(* IEC 61131-3 sources: TetherPLC/compat/tc2 (part 2) *)

(* ---- tc2_hvac.st ---- *)
// tc2_hvac.st — Tc2_HVAC surface (TF8000_TC3_HVAC_EN): pure-ST
// HVAC control blocks — no host/hardware dependency.  Covers
// the documented categories: actuators, motors/pumps, mux,
// redundancy, analog scaling, controllers (2-point, step, PID),
// sequence controllers, heating curve / outside-temp damping,
// alarm/anti-blocking/blink helpers, and BAR room-automation
// primitives.  Terminal bindings (KL32xx) are not modeled —
// the blocks operate on scaled process values.

// ---- FB_HVACAnalogInput: raw counts -> engineering value ----
FUNCTION_BLOCK FB_HVACAnalogInput
VAR_INPUT
    Raw : LREAL;                // raw counts
    RawMin : LREAL;
    RawMax : LREAL;
    EngMin : LREAL;
    EngMax : LREAL;
END_VAR
VAR_OUTPUT
    Value : LREAL;
END_VAR
    IF RawMax = RawMin THEN
        Value := EngMin;
    ELSE
        Value := EngMin + (Raw - RawMin) * (EngMax - EngMin) /
                 (RawMax - RawMin);
        IF Value < EngMin THEN Value := EngMin; END_IF;
        IF Value > EngMax THEN Value := EngMax; END_IF;
    END_IF;
END_FUNCTION_BLOCK

// ---- FB_HVACAnalogOutput: engineering value -> raw ----
FUNCTION_BLOCK FB_HVACAnalogOutput
VAR_INPUT
    Value : LREAL;
    EngMin : LREAL;
    EngMax : LREAL;
    RawMin : LREAL;
    RawMax : LREAL;
END_VAR
VAR_OUTPUT
    Raw : LREAL;
END_VAR
    IF EngMax = EngMin THEN
        Raw := RawMin;
    ELSE
        Raw := RawMin + (Value - EngMin) * (RawMax - RawMin) /
               (EngMax - EngMin);
        IF Raw < RawMin THEN Raw := RawMin; END_IF;
        IF Raw > RawMax THEN Raw := RawMax; END_IF;
    END_IF;
END_FUNCTION_BLOCK

// ---- FB_HVACScale: generic piecewise-linear scale ----
FUNCTION_BLOCK FB_HVACScale
VAR_INPUT
    x : LREAL;
    xMin : LREAL;
    xMax : LREAL;
    yMin : LREAL;
    yMax : LREAL;
END_VAR
VAR_OUTPUT
    y : LREAL;
END_VAR
    IF xMax = xMin THEN
        y := yMin;
    ELSE
        y := yMin + (x - xMin) * (yMax - yMin) / (xMax - xMin);
    END_IF;
END_FUNCTION_BLOCK

// ---- FB_HVAC2PointActuator: two-point damper/valve ----
// bCtrlVoltage TRUE -> run open; plus manual override and end-
// switch feedback monitoring.
FUNCTION_BLOCK FB_HVAC2PointActuator
VAR_INPUT
    bEnable : BOOL;
    bIn : BOOL;                 // demand: TRUE = open
    bManSwitch : BOOL;          // manual open override
    bLimitSwitchOpen : BOOL;
    bLimitSwitchClose : BOOL;
    tRun : LREAL;               // travel time s
    CycleTime : LREAL;
END_VAR
VAR_OUTPUT
    bOut : BOOL;                // drive command
    bFault : BOOL;              // end-switch disagreement
    Position : LREAL;           // 0 closed .. 100 open
END_VAR
VAR
    pos : LREAL;
END_VAR
    IF NOT bEnable THEN
        bOut := FALSE;
        bFault := FALSE;
        RETURN;
    END_IF;
    bOut := bIn OR bManSwitch;
    IF tRun > 0.0 THEN
        IF bOut THEN
            pos := pos + 100.0 * CycleTime / tRun;
            IF pos > 100.0 THEN pos := 100.0; END_IF;
        ELSE
            pos := pos - 100.0 * CycleTime / tRun;
            IF pos < 0.0 THEN pos := 0.0; END_IF;
        END_IF;
    END_IF;
    Position := pos;
    // fault: fully driven but feedback contradicts
    bFault := (pos >= 100.0 AND NOT bLimitSwitchOpen) OR
             (pos <= 0.0 AND NOT bLimitSwitchClose);
END_FUNCTION_BLOCK

// ---- FB_HVAC3PointActuator: three-point (open/close) ----
FUNCTION_BLOCK FB_HVAC3PointActuator
VAR_INPUT
    bEnable : BOOL;
    bOpen : BOOL;
    bClose : BOOL;
    tRun : LREAL;
    CycleTime : LREAL;
END_VAR
VAR_OUTPUT
    bOutOpen : BOOL;
    bOutClose : BOOL;
    Position : LREAL;
END_VAR
VAR
    pos : LREAL;
END_VAR
    IF NOT bEnable THEN
        bOutOpen := FALSE;
        bOutClose := FALSE;
        RETURN;
    END_IF;
    bOutOpen := bOpen AND NOT bClose;
    bOutClose := bClose AND NOT bOpen;
    IF tRun > 0.0 THEN
        IF bOutOpen THEN
            pos := pos + 100.0 * CycleTime / tRun;
            IF pos > 100.0 THEN pos := 100.0; END_IF;
        END_IF;
        IF bOutClose THEN
            pos := pos - 100.0 * CycleTime / tRun;
            IF pos < 0.0 THEN pos := 0.0; END_IF;
        END_IF;
    END_IF;
    Position := pos;
END_FUNCTION_BLOCK

// ---- FB_HVACCirculationPump: pump with standby lead swap ----
FUNCTION_BLOCK FB_HVACCirculationPump
VAR_INPUT
    bEnable : BOOL;
    bDemand : BOOL;
    bFault1 : BOOL;
    bFault2 : BOOL;
    bSwap : BOOL;               // lead-rotation request
END_VAR
VAR_OUTPUT
    bPump1 : BOOL;
    bPump2 : BOOL;
    Lead : INT;                 // 1 or 2
    bAlarm : BOOL;
END_VAR
VAR
    leadN : INT;
END_VAR
    IF leadN = 0 THEN leadN := 1; END_IF;
    IF bSwap THEN
        IF leadN = 1 THEN leadN := 2; ELSE leadN := 1; END_IF;
    END_IF;
    Lead := leadN;
    IF NOT bEnable OR NOT bDemand THEN
        bPump1 := FALSE;
        bPump2 := FALSE;
        bAlarm := bFault1 AND bFault2;
        RETURN;
    END_IF;
    bPump1 := leadN = 1 AND NOT bFault1;
    bPump2 := (leadN = 2 OR bFault1) AND NOT bFault2;
    bAlarm := bFault1 AND bFault2;
END_FUNCTION_BLOCK

// ---- FB_HVACMotor1Speed / Motor2Speed / Motor3Speed ----
FUNCTION_BLOCK FB_HVACMotor1Speed
VAR_INPUT
    bEnable : BOOL;
    Speed : INT;                // 0 off, 1 run
END_VAR
VAR_OUTPUT
    bOut1 : BOOL;
END_VAR
    bOut1 := bEnable AND Speed = 1;
END_FUNCTION_BLOCK

FUNCTION_BLOCK FB_HVACMotor2Speed
VAR_INPUT
    bEnable : BOOL;
    Speed : INT;                // 0..2
END_VAR
VAR_OUTPUT
    bOut1 : BOOL;
    bOut2 : BOOL;
END_VAR
    bOut1 := bEnable AND Speed = 1;
    bOut2 := bEnable AND Speed = 2;
END_FUNCTION_BLOCK

FUNCTION_BLOCK FB_HVACMotor3Speed
VAR_INPUT
    bEnable : BOOL;
    Speed : INT;                // 0..3
END_VAR
VAR_OUTPUT
    bOut1 : BOOL;
    bOut2 : BOOL;
    bOut3 : BOOL;
END_VAR
    bOut1 := bEnable AND Speed = 1;
    bOut2 := bEnable AND Speed = 2;
    bOut3 := bEnable AND Speed = 3;
END_FUNCTION_BLOCK

// ---- FB_HVACMux8: 8 -> 1 analog mux by selector ----
FUNCTION_BLOCK FB_HVACMux8
VAR_INPUT
    Sel : INT;                  // 1..8
    In1 : LREAL; In2 : LREAL; In3 : LREAL; In4 : LREAL;
    In5 : LREAL; In6 : LREAL; In7 : LREAL; In8 : LREAL;
END_VAR
VAR_OUTPUT
    Out : LREAL;
END_VAR
    IF Sel = 1 THEN Out := In1;
    ELSIF Sel = 2 THEN Out := In2;
    ELSIF Sel = 3 THEN Out := In3;
    ELSIF Sel = 4 THEN Out := In4;
    ELSIF Sel = 5 THEN Out := In5;
    ELSIF Sel = 6 THEN Out := In6;
    ELSIF Sel = 7 THEN Out := In7;
    ELSIF Sel = 8 THEN Out := In8;
    ELSE Out := 0.0;
    END_IF;
END_FUNCTION_BLOCK

// ---- FB_HVACMux8_BOOL: 8 -> 1 bool mux ----
FUNCTION_BLOCK FB_HVACMux8_BOOL
VAR_INPUT
    Sel : INT;
    In1 : BOOL; In2 : BOOL; In3 : BOOL; In4 : BOOL;
    In5 : BOOL; In6 : BOOL; In7 : BOOL; In8 : BOOL;
END_VAR
VAR_OUTPUT
    Out : BOOL;
END_VAR
    IF Sel = 1 THEN Out := In1;
    ELSIF Sel = 2 THEN Out := In2;
    ELSIF Sel = 3 THEN Out := In3;
    ELSIF Sel = 4 THEN Out := In4;
    ELSIF Sel = 5 THEN Out := In5;
    ELSIF Sel = 6 THEN Out := In6;
    ELSIF Sel = 7 THEN Out := In7;
    ELSIF Sel = 8 THEN Out := In8;
    ELSE Out := FALSE;
    END_IF;
END_FUNCTION_BLOCK

// ---- FB_HVACRedundancyCtrl: n+1 pump/fan redundancy ----
// N units, need Required running; rotates the lead and covers
// faults in order.
FUNCTION_BLOCK FB_HVACRedundancyCtrl
VAR_INPUT
    bEnable : BOOL;
    Required : INT;             // units demanded 0..3
    bFault1 : BOOL;
    bFault2 : BOOL;
    bFault3 : BOOL;
    bRotate : BOOL;
END_VAR
VAR_OUTPUT
    bOut1 : BOOL;
    bOut2 : BOOL;
    bOut3 : BOOL;
    Lead : INT;
    bAlarm : BOOL;
END_VAR
VAR
    leadN : INT;
    want : INT;
    ok1 : BOOL;
    ok2 : BOOL;
    ok3 : BOOL;
END_VAR
    IF leadN = 0 THEN leadN := 1; END_IF;
    IF bRotate THEN
        leadN := leadN + 1;
        IF leadN > 3 THEN leadN := 1; END_IF;
    END_IF;
    Lead := leadN;
    ok1 := NOT bFault1;
    ok2 := NOT bFault2;
    ok3 := NOT bFault3;
    want := Required;
    bOut1 := FALSE; bOut2 := FALSE; bOut3 := FALSE;
    IF bEnable THEN
        // start at leadN, wrap, pick healthy units
        IF want > 0 THEN
            IF leadN = 1 THEN
                IF ok1 THEN bOut1 := TRUE; want := want - 1; END_IF;
                IF want > 0 AND ok2 THEN bOut2 := TRUE; want := want - 1; END_IF;
                IF want > 0 AND ok3 THEN bOut3 := TRUE; want := want - 1; END_IF;
            ELSIF leadN = 2 THEN
                IF ok2 THEN bOut2 := TRUE; want := want - 1; END_IF;
                IF want > 0 AND ok3 THEN bOut3 := TRUE; want := want - 1; END_IF;
                IF want > 0 AND ok1 THEN bOut1 := TRUE; want := want - 1; END_IF;
            ELSE
                IF ok3 THEN bOut3 := TRUE; want := want - 1; END_IF;
                IF want > 0 AND ok1 THEN bOut1 := TRUE; want := want - 1; END_IF;
                IF want > 0 AND ok2 THEN bOut2 := TRUE; want := want - 1; END_IF;
            END_IF;
        END_IF;
    END_IF;
    bAlarm := want > 0;         // couldn't satisfy demand
END_FUNCTION_BLOCK

// ---- FB_HVAC2PointCtrl: on/off controller with hysteresis ----
FUNCTION_BLOCK FB_HVAC2PointCtrl
VAR_INPUT
    bEnable : BOOL;
    fActual : LREAL;
    fSetpoint : LREAL;
    fHysteresis : LREAL;
    bInvert : BOOL;             // TRUE = cooling (on above SP)
END_VAR
VAR_OUTPUT
    bOut : BOOL;
END_VAR
VAR
    q : BOOL;
END_VAR
    IF NOT bEnable THEN q := FALSE; bOut := FALSE; RETURN; END_IF;
    IF bInvert THEN
        IF fActual >= fSetpoint + fHysteresis THEN q := TRUE; END_IF;
        IF fActual <= fSetpoint THEN q := FALSE; END_IF;
    ELSE
        IF fActual <= fSetpoint - fHysteresis THEN q := TRUE; END_IF;
        IF fActual >= fSetpoint THEN q := FALSE; END_IF;
    END_IF;
    bOut := q;
END_FUNCTION_BLOCK

// ---- FB_HVACI_CtrlStep: staged step controller ----
// Splits the control error into up to 4 equal stages.
FUNCTION_BLOCK FB_HVACI_CtrlStep
VAR_INPUT
    bEnable : BOOL;
    fActual : LREAL;
    fSetpoint : LREAL;
    fStepRange : LREAL;         // error span for all 4 stages
    nStages : INT;              // 1..4
END_VAR
VAR_OUTPUT
    bStage1 : BOOL;
    bStage2 : BOOL;
    bStage3 : BOOL;
    bStage4 : BOOL;
END_VAR
VAR
    e : LREAL;
    step : LREAL;
END_VAR
    IF NOT bEnable OR nStages <= 0 OR fStepRange <= 0.0 THEN
        bStage1 := FALSE; bStage2 := FALSE;
        bStage3 := FALSE; bStage4 := FALSE;
        RETURN;
    END_IF;
    e := fSetpoint - fActual;
    step := fStepRange / DINT_TO_LREAL(INT_TO_DINT(nStages));
    bStage1 := e >= step;
    bStage2 := nStages >= 2 AND e >= 2.0 * step;
    bStage3 := nStages >= 3 AND e >= 3.0 * step;
    bStage4 := nStages >= 4 AND e >= 4.0 * step;
END_FUNCTION_BLOCK

// ---- FB_HVACPIDCtrl: PI(D) controller ----
// Incremental PID with anti-windup clamp on the output.
FUNCTION_BLOCK FB_HVACPIDCtrl
VAR_INPUT
    bEnable : BOOL;
    fActual : LREAL;
    fSetpoint : LREAL;
    fKp : LREAL;
    fTi : LREAL;                // s; 0 = P only
    fTd : LREAL;                // s
    fOutMin : LREAL;
    fOutMax : LREAL;
    CycleTime : LREAL;
END_VAR
VAR_OUTPUT
    fOut : LREAL;
    fError : LREAL;
END_VAR
VAR
    iTerm : LREAL;
    ePrev : LREAL;
END_VAR
    IF NOT bEnable THEN
        fOut := fOutMin;
        iTerm := 0.0;
        ePrev := 0.0;
        fError := 0.0;
        RETURN;
    END_IF;
    fError := fSetpoint - fActual;
    iTerm := iTerm + fError * CycleTime;
    fOut := fKp * (fError + ePrev);
    IF fTi > 0.0 THEN
        fOut := fKp * (fError + iTerm / fTi);
    END_IF;
    IF fTd > 0.0 AND CycleTime > 0.0 THEN
        fOut := fOut + fKp * fTd * (fError - ePrev) / CycleTime;
    END_IF;
    IF fOut > fOutMax THEN
        fOut := fOutMax;
        iTerm := iTerm - fError * CycleTime;   // anti-windup
    END_IF;
    IF fOut < fOutMin THEN
        fOut := fOutMin;
        iTerm := iTerm - fError * CycleTime;
    END_IF;
    ePrev := fError;
END_FUNCTION_BLOCK

// ---- FB_HVACHeatingCurve: outdoor-reset flow setpoint ----
// Flow SP = fSpMin + (fSpMax-fSpMin) * (tRoom - tOut) /
// (tRoom - tOutMin) when outside is cold, clamped.
FUNCTION_BLOCK FB_HVACHeatingCurve
VAR_INPUT
    bEnable : BOOL;
    fOutsideTemp : LREAL;
    fOutsideMin : LREAL;        // design outside temp
    fRoomTemp : LREAL;
    fSpMin : LREAL;             // flow SP at warm extreme
    fSpMax : LREAL;             // flow SP at design outside
END_VAR
VAR_OUTPUT
    fFlowSp : LREAL;
END_VAR
    IF NOT bEnable OR fRoomTemp = fOutsideMin THEN
        fFlowSp := fSpMin;
        RETURN;
    END_IF;
    fFlowSp := fSpMin + (fSpMax - fSpMin) *
               (fRoomTemp - fOutsideTemp) / (fRoomTemp - fOutsideMin);
    IF fFlowSp > fSpMax THEN fFlowSp := fSpMax; END_IF;
    IF fFlowSp < fSpMin THEN fFlowSp := fSpMin; END_IF;
END_FUNCTION_BLOCK

// ---- FB_HVACOutsideTempDamped: damped outdoor temperature ----
// First-order lag on the measured outside temperature.
FUNCTION_BLOCK FB_HVACOutsideTempDamped
VAR_INPUT
    bEnable : BOOL;
    fOutsideTemp : LREAL;
    fTau : LREAL;               // damping time constant s
    CycleTime : LREAL;
END_VAR
VAR_OUTPUT
    fDamped : LREAL;
END_VAR
VAR
    y : LREAL;
    init : BOOL;
END_VAR
    IF NOT bEnable THEN
        init := FALSE;
        RETURN;
    END_IF;
    IF NOT init OR fTau <= 0.0 THEN
        y := fOutsideTemp;
        init := TRUE;
    ELSE
        y := y + (fOutsideTemp - y) * CycleTime / fTau;
    END_IF;
    fDamped := y;
END_FUNCTION_BLOCK

// ---- FB_HVACSetpointRamp: ramp a setpoint to target ----
FUNCTION_BLOCK FB_HVACSetpointRamp
VAR_INPUT
    bEnable : BOOL;
    fTarget : LREAL;
    fSlew : LREAL;              // unit/s
    CycleTime : LREAL;
END_VAR
VAR_OUTPUT
    fOut : LREAL;
    bDone : BOOL;
END_VAR
    IF NOT bEnable THEN bDone := FALSE; RETURN; END_IF;
    IF fOut < fTarget THEN
        fOut := fOut + fSlew * CycleTime;
        IF fOut > fTarget THEN fOut := fTarget; END_IF;
    ELSIF fOut > fTarget THEN
        fOut := fOut - fSlew * CycleTime;
        IF fOut < fTarget THEN fOut := fTarget; END_IF;
    END_IF;
    bDone := fOut = fTarget;
END_FUNCTION_BLOCK

// ---- FB_HVACAlarm: limit alarm with hysteresis + delay ----
FUNCTION_BLOCK FB_HVACAlarm
VAR_INPUT
    bEnable : BOOL;
    fValue : LREAL;
    fLimit : LREAL;
    fHysteresis : LREAL;
    tDelay : LREAL;             // s before alarm latches
    bAck : BOOL;
    CycleTime : LREAL;
END_VAR
VAR_OUTPUT
    bAlarm : BOOL;
    bActive : BOOL;             // condition currently true
END_VAR
VAR
    tAcc : LREAL;
    latch : BOOL;
END_VAR
    IF NOT bEnable THEN
        bAlarm := FALSE; bActive := FALSE; latch := FALSE;
        tAcc := 0.0;
        RETURN;
    END_IF;
    bActive := fValue >= fLimit;
    IF bActive THEN
        tAcc := tAcc + CycleTime;
        IF tAcc >= tDelay THEN latch := TRUE; END_IF;
    END_IF;
    IF fValue <= fLimit - fHysteresis THEN tAcc := 0.0; END_IF;
    IF bAck THEN latch := FALSE; END_IF;
    bAlarm := latch;
END_FUNCTION_BLOCK

// ---- FB_HVACAntiBlockingPump: periodic exercise run ----
// If the pump has been idle longer than tIdle, run it for
// tRunTime to prevent seizing.
FUNCTION_BLOCK FB_HVACAntiBlockingPump
VAR_INPUT
    bEnable : BOOL;
    bDemand : BOOL;
    tIdle : LREAL;              // s idle before exercise
    tRunTime : LREAL;           // s exercise duration
    CycleTime : LREAL;
END_VAR
VAR_OUTPUT
    bPump : BOOL;
    bExercise : BOOL;           // exercising (not demand)
END_VAR
VAR
    tIdleAcc : LREAL;
    tRunAcc : LREAL;
END_VAR
    IF NOT bEnable THEN
        bPump := FALSE; bExercise := FALSE;
        tIdleAcc := 0.0; tRunAcc := 0.0;
        RETURN;
    END_IF;
    IF bDemand THEN
        tIdleAcc := 0.0;
        tRunAcc := 0.0;
        bPump := TRUE;
        bExercise := FALSE;
    ELSIF tRunAcc > 0.0 THEN
        tRunAcc := tRunAcc - CycleTime;
        bPump := tRunAcc > 0.0;
        bExercise := bPump;
        IF NOT bExercise THEN tIdleAcc := 0.0; END_IF;
    ELSE
        tIdleAcc := tIdleAcc + CycleTime;
        IF tIdleAcc >= tIdle THEN
            tRunAcc := tRunTime;
            tIdleAcc := 0.0;
        END_IF;
        bPump := FALSE;
        bExercise := FALSE;
    END_IF;
END_FUNCTION_BLOCK

// ---- FB_HVACBlink: square-wave blinker ----
FUNCTION_BLOCK FB_HVACBlink
VAR_INPUT
    bEnable : BOOL;
    tOn : LREAL;                // s
    tOff : LREAL;               // s
    CycleTime : LREAL;
END_VAR
VAR_OUTPUT
    bOut : BOOL;
END_VAR
VAR
    tAcc : LREAL;
    q : BOOL;
END_VAR
    IF NOT bEnable THEN bOut := FALSE; q := FALSE; tAcc := 0.0; RETURN; END_IF;
    tAcc := tAcc + CycleTime;
    IF q THEN
        IF tAcc >= tOn THEN q := FALSE; tAcc := 0.0; END_IF;
    ELSE
        IF tAcc >= tOff THEN q := TRUE; tAcc := 0.0; END_IF;
    END_IF;
    bOut := q;
END_FUNCTION_BLOCK

// ---- FB_HVACPIDHeating / Cooling convenience wrappers ----
// Sequence controllers in the catalogue are PID + mode glue;
// the core PID is FB_HVACPIDCtrl above.

// ---- FB_BARSetpointRoom: room setpoint with shift ----
FUNCTION_BLOCK FB_BARSetpointRoom
VAR_INPUT
    bEnable : BOOL;
    fBaseSp : LREAL;            // base comfort setpoint
    fShift : LREAL;             // user shift +-K
    fShiftMax : LREAL;
END_VAR
VAR_OUTPUT
    fSetpoint : LREAL;
END_VAR
    IF NOT bEnable THEN fSetpoint := fBaseSp; RETURN; END_IF;
    fSetpoint := fBaseSp + fShift;
    IF fSetpoint > fBaseSp + fShiftMax THEN
        fSetpoint := fBaseSp + fShiftMax;
    END_IF;
    IF fSetpoint < fBaseSp - fShiftMax THEN
        fSetpoint := fBaseSp - fShiftMax;
    END_IF;
END_FUNCTION_BLOCK

// ---- FB_BARDelayedHysteresis: on/off delay on a level ----
FUNCTION_BLOCK FB_BARDelayedHysteresis
VAR_INPUT
    bEnable : BOOL;
    fValue : LREAL;
    fOn : LREAL;
    fOff : LREAL;
    tOnDelay : LREAL;
    tOffDelay : LREAL;
    CycleTime : LREAL;
END_VAR
VAR_OUTPUT
    bOut : BOOL;
END_VAR
VAR
    tAcc : LREAL;
    q : BOOL;
END_VAR
    IF NOT bEnable THEN bOut := FALSE; q := FALSE; tAcc := 0.0; RETURN; END_IF;
    IF fValue >= fOn AND NOT q THEN
        tAcc := tAcc + CycleTime;
        IF tAcc >= tOnDelay THEN q := TRUE; tAcc := 0.0; END_IF;
    ELSIF fValue <= fOff AND q THEN
        tAcc := tAcc + CycleTime;
        IF tAcc >= tOffDelay THEN q := FALSE; tAcc := 0.0; END_IF;
    ELSE
        tAcc := 0.0;
    END_IF;
    bOut := q;
END_FUNCTION_BLOCK

(* ---- tc2_iec61850.st ---- *)
// tc2_iec61850.st — TwinCAT IEC 61850 client surface (Tc3_IEC61850 /
// TF6101 shape) over the tplc-iec61850 service + FB_Iec61850 builtin.
//
// The PLC is the client (control-center side) over the full OSI
// stack via libiec61850: FB_Iec61850Connect runs TPKT/COTP/Session/
// Presentation/ACSE/MMS Initiate; FB_Iec61850Read/Write carry
// Confirmed-Request Read/Write on domain+item named variables;
// FB_Iec61850GetNameList lists a domain's objects; Disconnect
// releases.  Reporting/RCB, GOOSE/SMV, and the full data model are
// out of scope for this tranche.
//
// Object addressing is a domain (Logical Device) name + an item
// (VariableAccess) name — "tetherTestLD" + "LLN0$Health$stVal".
// Values travel as bounded STRING[255] (numerics as ASCII repr,
// structured values as their MmsValue string).  STATUS carries the
// service return code, ErrorID its positive form + the last MMS
// service error via FB_Iec61850Status.

// ---- FB_Iec61850Connect: TCP + OSI associate + MMS Initiate ----
FUNCTION_BLOCK FB_Iec61850Connect
VAR_INPUT
    Execute : BOOL;
    RemoteHost : STRING[63];
    RemotePort : UDINT;
END_VAR
VAR_OUTPUT
    Done : BOOL;
    Busy : BOOL;
    Error : BOOL;
    ErrorID : UDINT;
    ConnectionHdl : UDINT;
END_VAR
VAR
    ch : FB_Iec61850;
    exPrev : BOOL;
END_VAR
    Done := FALSE;
    Error := FALSE;
    ErrorID := 0;
    IF Execute AND NOT exPrev THEN
        ch.OP := 1;
        ch.HOST := RemoteHost;
        ch.PORT := RemotePort;
        ch();
        IF ch.STATUS = 0 THEN
            Done := TRUE;
            ConnectionHdl := ch.HANDLE;
        ELSE
            Error := TRUE;
            ErrorID := ch.ERRID;
        END_IF;
    END_IF;
    exPrev := Execute;
    Busy := FALSE;
END_FUNCTION_BLOCK

// ---- FB_Iec61850Disconnect: release the association ----
FUNCTION_BLOCK FB_Iec61850Disconnect
VAR_INPUT
    Execute : BOOL;
    ConnectionHdl : UDINT;
END_VAR
VAR_OUTPUT
    Done : BOOL;
    Busy : BOOL;
    Error : BOOL;
    ErrorID : UDINT;
END_VAR
VAR
    ch : FB_Iec61850;
    exPrev : BOOL;
END_VAR
    Done := FALSE;
    Error := FALSE;
    ErrorID := 0;
    IF Execute AND NOT exPrev THEN
        ch.OP := 2;
        ch.HANDLE := ConnectionHdl;
        ch();
        IF ch.STATUS = 0 THEN
            Done := TRUE;
        ELSE
            Error := TRUE;
            ErrorID := ch.ERRID;
        END_IF;
    END_IF;
    exPrev := Execute;
    Busy := FALSE;
END_FUNCTION_BLOCK

// ---- FB_Iec61850Status: association status ----
FUNCTION_BLOCK FB_Iec61850Status
VAR_INPUT
    Execute : BOOL;
    ConnectionHdl : UDINT;
END_VAR
VAR_OUTPUT
    Done : BOOL;
    Error : BOOL;
    ErrorID : UDINT;
    ConnectionState : DINT;
    InvokeId : UDINT;
    LastMmsError : UDINT;
END_VAR
VAR
    ch : FB_Iec61850;
END_VAR
    Done := FALSE;
    Error := FALSE;
    ErrorID := 0;
    IF Execute THEN
        ch.OP := 3;
        ch.HANDLE := ConnectionHdl;
        ch();
        IF ch.STATUS = 0 THEN
            Done := TRUE;
            ConnectionState := ch.STATE;
            InvokeId := ch.INVOKE;
            LastMmsError := ch.LASTERR;
        ELSE
            Error := TRUE;
            ErrorID := ch.ERRID;
        END_IF;
    END_IF;
END_FUNCTION_BLOCK

// ---- FB_Iec61850Read: Confirmed-Request Read ----
FUNCTION_BLOCK FB_Iec61850Read
VAR_INPUT
    Execute : BOOL;
    ConnectionHdl : UDINT;
    Domain : STRING[63];
    Item : STRING[127];
END_VAR
VAR_OUTPUT
    Done : BOOL;
    Error : BOOL;
    ErrorID : UDINT;
    Value : STRING[255];
END_VAR
VAR
    ch : FB_Iec61850;
    exPrev : BOOL;
END_VAR
    Done := FALSE;
    Error := FALSE;
    ErrorID := 0;
    IF Execute AND NOT exPrev THEN
        ch.OP := 4;
        ch.HANDLE := ConnectionHdl;
        ch.DOMAIN := Domain;
        ch.ITEM := Item;
        ch();
        IF ch.STATUS >= 0 THEN
            Done := TRUE;
            Value := ch.VAL;
        ELSE
            Error := TRUE;
            ErrorID := ch.ERRID;
        END_IF;
    END_IF;
    exPrev := Execute;
END_FUNCTION_BLOCK

// ---- FB_Iec61850Write: Confirmed-Request Write ----
FUNCTION_BLOCK FB_Iec61850Write
VAR_INPUT
    Execute : BOOL;
    ConnectionHdl : UDINT;
    Domain : STRING[63];
    Item : STRING[127];
    Value : STRING[255];
END_VAR
VAR_OUTPUT
    Done : BOOL;
    Error : BOOL;
    ErrorID : UDINT;
END_VAR
VAR
    ch : FB_Iec61850;
    exPrev : BOOL;
END_VAR
    Done := FALSE;
    Error := FALSE;
    ErrorID := 0;
    IF Execute AND NOT exPrev THEN
        ch.OP := 5;
        ch.HANDLE := ConnectionHdl;
        ch.DOMAIN := Domain;
        ch.ITEM := Item;
        ch.VAL := Value;
        ch();
        IF ch.STATUS = 0 THEN
            Done := TRUE;
        ELSE
            Error := TRUE;
            ErrorID := ch.ERRID;
        END_IF;
    END_IF;
    exPrev := Execute;
END_FUNCTION_BLOCK

// ---- FB_Iec61850GetNameList: MMS GetNameList on a domain ----
FUNCTION_BLOCK FB_Iec61850GetNameList
VAR_INPUT
    Execute : BOOL;
    ConnectionHdl : UDINT;
    Domain : STRING[63];
END_VAR
VAR_OUTPUT
    Done : BOOL;
    Error : BOOL;
    ErrorID : UDINT;
    NameList : STRING[255];
END_VAR
VAR
    ch : FB_Iec61850;
    exPrev : BOOL;
END_VAR
    Done := FALSE;
    Error := FALSE;
    ErrorID := 0;
    IF Execute AND NOT exPrev THEN
        ch.OP := 6;
        ch.HANDLE := ConnectionHdl;
        ch.DOMAIN := Domain;
        ch();
        IF ch.STATUS >= 0 THEN
            Done := TRUE;
            NameList := ch.VAL;
        ELSE
            Error := TRUE;
            ErrorID := ch.ERRID;
        END_IF;
    END_IF;
    exPrev := Execute;
END_FUNCTION_BLOCK

// ---- FB_Iec61850RCBGet: MMS GetRCBValues on an RCB reference ----
// RcbRef is the MMS object reference of the report control block,
// e.g. 'tetherIEDtetherTestLD/LLN0$BR$MeasURCB'.
FUNCTION_BLOCK FB_Iec61850RCBGet
VAR_INPUT
    Execute : BOOL;
    ConnectionHdl : UDINT;
    RcbRef : STRING[127];
END_VAR
VAR_OUTPUT
    Done : BOOL;
    Error : BOOL;
    ErrorID : UDINT;
    RptId : STRING[31];
    DataSet : STRING[63];
    ConfRev : UDINT;
    BufTm : UDINT;
    IntgPd : UDINT;
    SqNum : UDINT;
    OptFlds : UDINT;
    TrgOps : UDINT;
    RptEna : BOOL;
    Resv : BOOL;
    Buffered : BOOL;
    GI : BOOL;
    PurgeBuf : BOOL;
    ResvTms : UDINT;
    EntryId : UDINT;
END_VAR
VAR
    ch : FB_Iec61850;
    exPrev : BOOL;
END_VAR
    Done := FALSE;
    Error := FALSE;
    ErrorID := 0;
    IF Execute AND NOT exPrev THEN
        ch.OP := 7;
        ch.HANDLE := ConnectionHdl;
        ch.RCBREF := RcbRef;
        ch();
        IF ch.STATUS = 0 THEN
            Done := TRUE;
            RptId := ch.RPTID;
            DataSet := ch.DATASET;
            ConfRev := ch.CONFREV;
            BufTm := ch.BUFTM;
            IntgPd := ch.INTGPD;
            SqNum := ch.SQNUM;
            OptFlds := ch.OPTFLDS;
            TrgOps := ch.TRGOPS;
            RptEna := ch.RPTENA <> 0;
            Resv := ch.RESV <> 0;
            Buffered := ch.BUFFERED <> 0;
            GI := ch.GI <> 0;
            PurgeBuf := ch.PURGEBUF <> 0;
            ResvTms := ch.RESVTMS;
            EntryId := ch.ENTRYID;
        ELSE
            Error := TRUE;
            ErrorID := ch.ERRID;
        END_IF;
    END_IF;
    exPrev := Execute;
END_FUNCTION_BLOCK

// ---- FB_Iec61850RCBSet: MMS SetRCBValues (URCB-safe subset) ----
// Flags: bit0 RptEna, bit1 Resv, bit2 GI, bit3 PurgeBuf (buffered
// RCBs only).  Once the RCB is enabled the service narrows the write
// to the attributes servers accept in that state (RptEna disable,
// GI, PurgeBuf); a redundant enable is a no-op.  Enabling installs
// the report handler on the connection.
FUNCTION_BLOCK FB_Iec61850RCBSet
VAR_INPUT
    Execute : BOOL;
    ConnectionHdl : UDINT;
    RcbRef : STRING[127];
    Flags : UDINT;
END_VAR
VAR_OUTPUT
    Done : BOOL;
    Error : BOOL;
    ErrorID : UDINT;
END_VAR
VAR
    ch : FB_Iec61850;
    exPrev : BOOL;
END_VAR
    Done := FALSE;
    Error := FALSE;
    ErrorID := 0;
    IF Execute AND NOT exPrev THEN
        ch.OP := 8;
        ch.HANDLE := ConnectionHdl;
        ch.RCBREF := RcbRef;
        ch.FLAGS := Flags;
        ch();
        IF ch.STATUS = 0 THEN
            Done := TRUE;
        ELSE
            Error := TRUE;
            ErrorID := ch.ERRID;
        END_IF;
    END_IF;
    exPrev := Execute;
END_FUNCTION_BLOCK

// ---- FB_Iec61850ReportPoll: drain received reports ----
// Report holds newline-separated "dataset|v0,v1,..." lines received
// since the last poll; ReportBytes is the drained byte count.
FUNCTION_BLOCK FB_Iec61850ReportPoll
VAR_INPUT
    Execute : BOOL;
    ConnectionHdl : UDINT;
END_VAR
VAR_OUTPUT
    Done : BOOL;
    Error : BOOL;
    ErrorID : UDINT;
    Report : STRING[255];
    ReportBytes : UDINT;
END_VAR
VAR
    ch : FB_Iec61850;
    exPrev : BOOL;
END_VAR
    Done := FALSE;
    Error := FALSE;
    ErrorID := 0;
    Report := '';
    ReportBytes := 0;
    IF Execute AND NOT exPrev THEN
        ch.OP := 9;
        ch.HANDLE := ConnectionHdl;
        ch();
        IF ch.STATUS >= 0 THEN
            Done := TRUE;
            Report := ch.VAL;
            ReportBytes := ch.RCNT;
        ELSE
            Error := TRUE;
            ErrorID := ch.ERRID;
        END_IF;
    END_IF;
    exPrev := Execute;
END_FUNCTION_BLOCK

// ---- FB_Iec61850Control: controllable data object command ----
// ObjectRef is the "domain/LN.DO" reference (e.g.
// "tetherTestLD/LLN0.SWI1").  Mode: 1=Select, 2=SelectWithValue,
// 3=Operate, 4=Cancel.  CtlValue is the ASCII control value
// ("true"/"false", integer or float text) for SelectWithValue and
// Operate.  Command termination arrives asynchronously — poll it
// with FB_Iec61850ControlPoll.
FUNCTION_BLOCK FB_Iec61850Control
VAR_INPUT
    Execute : BOOL;
    ConnectionHdl : UDINT;
    ObjectRef : STRING[127];
    Mode : UDINT;
    CtlValue : STRING[63];
END_VAR
VAR_OUTPUT
    Done : BOOL;
    Error : BOOL;
    ErrorID : UDINT;
    Value : STRING[63];
END_VAR
VAR
    ch : FB_Iec61850;
    exPrev : BOOL;
END_VAR
    Done := FALSE;
    Error := FALSE;
    ErrorID := 0;
    Value := '';
    IF Execute AND NOT exPrev THEN
        ch.OP := 10;
        ch.HANDLE := ConnectionHdl;
        ch.CTRLREF := ObjectRef;
        ch.CMODE := Mode;
        ch.CTLVAL := CtlValue;
        ch();
        IF ch.STATUS >= 0 THEN
            Done := TRUE;
            Value := ch.VAL;
        ELSE
            Error := TRUE;
            ErrorID := ch.ERRID;
        END_IF;
    END_IF;
    exPrev := Execute;
END_FUNCTION_BLOCK

// ---- FB_Iec61850ControlPoll: drain a CommandTermination event ----
// Pending is TRUE when an event was returned: Success marks
// CommandTermination+ vs -, Type is 0=select 1=operate 2=cancel,
// CtlNum echoes the server's control number.
FUNCTION_BLOCK FB_Iec61850ControlPoll
VAR_INPUT
    Execute : BOOL;
    ConnectionHdl : UDINT;
END_VAR
VAR_OUTPUT
    Done : BOOL;
    Error : BOOL;
    ErrorID : UDINT;
    Pending : BOOL;
    InvokeID : UDINT;
    Success : BOOL;
    Err : UDINT;
    EvType : UDINT;
    CtlNum : UDINT;
END_VAR
VAR
    ch : FB_Iec61850;
    exPrev : BOOL;
END_VAR
    Done := FALSE;
    Error := FALSE;
    ErrorID := 0;
    Pending := FALSE;
    InvokeID := 0;
    Success := FALSE;
    Err := 0;
    EvType := 0;
    CtlNum := 0;
    IF Execute AND NOT exPrev THEN
        ch.OP := 11;
        ch.HANDLE := ConnectionHdl;
        ch();
        IF ch.STATUS >= 0 THEN
            Done := TRUE;
            Pending := ch.CTLPEND > 0;
            InvokeID := ch.CTLINVOKE;
            Success := ch.CTLSUCCESS > 0;
            Err := ch.CTLERR;
            EvType := ch.CTLTYPE;
            CtlNum := ch.CTLNUM;
        ELSE
            Error := TRUE;
            ErrorID := ch.ERRID;
        END_IF;
    END_IF;
    exPrev := Execute;
END_FUNCTION_BLOCK

// ---- FB_Iec61850DataSetRead: MMS ReadDataSet ----
// DataSetRef is the MMS object reference of the data set, e.g.
// 'tetherIEDtetherTestLD/LLN0.measds' ('@name' for VMD scope).
// Values holds newline-separated "FCDA=value" lines; ElementCount
// is the number of data set members returned.
FUNCTION_BLOCK FB_Iec61850DataSetRead
VAR_INPUT
    Execute : BOOL;
    ConnectionHdl : UDINT;
    DataSetRef : STRING[127];
END_VAR
VAR_OUTPUT
    Done : BOOL;
    Error : BOOL;
    ErrorID : UDINT;
    Values : STRING[255];
    ElementCount : UDINT;
END_VAR
VAR
    ch : FB_Iec61850;
    exPrev : BOOL;
END_VAR
    Done := FALSE;
    Error := FALSE;
    ErrorID := 0;
    Values := '';
    ElementCount := 0;
    IF Execute AND NOT exPrev THEN
        ch.OP := 12;
        ch.HANDLE := ConnectionHdl;
        ch.DSREF := DataSetRef;
        ch();
        IF ch.STATUS >= 0 THEN
            Done := TRUE;
            Values := ch.VAL;
            ElementCount := ch.DSCOUNT;
        ELSE
            Error := TRUE;
            ErrorID := ch.ERRID;
        END_IF;
    END_IF;
    exPrev := Execute;
END_FUNCTION_BLOCK

// ---- FB_Iec61850DataSetDirectory: MMS GetDataSetDirectory ----
// Names holds the newline-separated FCDA object references of the
// data set members (same order as ReadDataSet values).
FUNCTION_BLOCK FB_Iec61850DataSetDirectory
VAR_INPUT
    Execute : BOOL;
    ConnectionHdl : UDINT;
    DataSetRef : STRING[127];
END_VAR
VAR_OUTPUT
    Done : BOOL;
    Error : BOOL;
    ErrorID : UDINT;
    Names : STRING[255];
    ElementCount : UDINT;
END_VAR
VAR
    ch : FB_Iec61850;
    exPrev : BOOL;
END_VAR
    Done := FALSE;
    Error := FALSE;
    ErrorID := 0;
    Names := '';
    ElementCount := 0;
    IF Execute AND NOT exPrev THEN
        ch.OP := 13;
        ch.HANDLE := ConnectionHdl;
        ch.DSREF := DataSetRef;
        ch();
        IF ch.STATUS >= 0 THEN
            Done := TRUE;
            Names := ch.VAL;
            ElementCount := ch.DSCOUNT;
        ELSE
            Error := TRUE;
            ErrorID := ch.ERRID;
        END_IF;
    END_IF;
    exPrev := Execute;
END_FUNCTION_BLOCK

// ---- FB_Iec61850DataSetWrite: MMS WriteDataSet ----
// Values is the same newline-separated shape ReadDataSet produces
// ("FCDA=value" lines or bare values in member order); member
// types come from a fresh ReadDataSet on the server.
FUNCTION_BLOCK FB_Iec61850DataSetWrite
VAR_INPUT
    Execute : BOOL;
    ConnectionHdl : UDINT;
    DataSetRef : STRING[127];
    Values : STRING[255];
END_VAR
VAR_OUTPUT
    Done : BOOL;
    Error : BOOL;
    ErrorID : UDINT;
END_VAR
VAR
    ch : FB_Iec61850;
    exPrev : BOOL;
END_VAR
    Done := FALSE;
    Error := FALSE;
    ErrorID := 0;
    IF Execute AND NOT exPrev THEN
        ch.OP := 14;
        ch.HANDLE := ConnectionHdl;
        ch.DSREF := DataSetRef;
        ch.VAL := Values;
        ch();
        IF ch.STATUS = 0 THEN
            Done := TRUE;
        ELSE
            Error := TRUE;
            ErrorID := ch.ERRID;
        END_IF;
    END_IF;
    exPrev := Execute;
END_FUNCTION_BLOCK

// ---- FB_Iec61850DataSetCreate: MMS CreateDataSet ----
// Elements is a newline-separated list of FCDA object references
// ("LD/LN.item[FC]" lines) defining the members.  DataSetRef uses the
// "LD/LN.name" form or "@name" for an association-specific set.
FUNCTION_BLOCK FB_Iec61850DataSetCreate
VAR_INPUT
    Execute : BOOL;
    ConnectionHdl : UDINT;
    DataSetRef : STRING[127];
    Elements : STRING[255];
END_VAR
VAR_OUTPUT
    Done : BOOL;
    Error : BOOL;
    ErrorID : UDINT;
END_VAR
VAR
    ch : FB_Iec61850;
    exPrev : BOOL;
END_VAR
    Done := FALSE;
    Error := FALSE;
    ErrorID := 0;
    IF Execute AND NOT exPrev THEN
        ch.OP := 15;
        ch.HANDLE := ConnectionHdl;
        ch.DSREF := DataSetRef;
        ch.VAL := Elements;
        ch();
        IF ch.STATUS = 0 THEN
            Done := TRUE;
        ELSE
            Error := TRUE;
            ErrorID := ch.ERRID;
        END_IF;
    END_IF;
    exPrev := Execute;
END_FUNCTION_BLOCK

// ---- FB_Iec61850DataSetDelete: MMS DeleteDataSet ----
FUNCTION_BLOCK FB_Iec61850DataSetDelete
VAR_INPUT
    Execute : BOOL;
    ConnectionHdl : UDINT;
    DataSetRef : STRING[127];
END_VAR
VAR_OUTPUT
    Done : BOOL;
    Error : BOOL;
    ErrorID : UDINT;
END_VAR
VAR
    ch : FB_Iec61850;
    exPrev : BOOL;
END_VAR
    Done := FALSE;
    Error := FALSE;
    ErrorID := 0;
    IF Execute AND NOT exPrev THEN
        ch.OP := 16;
        ch.HANDLE := ConnectionHdl;
        ch.DSREF := DataSetRef;
        ch();
        IF ch.STATUS = 0 THEN
            Done := TRUE;
        ELSE
            Error := TRUE;
            ErrorID := ch.ERRID;
        END_IF;
    END_IF;
    exPrev := Execute;
END_FUNCTION_BLOCK

(* ---- tc2_iofunctions.st ---- *)
// Tc2_IoFunctions -> general I/O enumeration surface.
// The 81-entry library is mostly EtherCAT device profiles (ASi,
// Profibus DPV1, Lightbus, CANopen, RAID, ...).  Those need the
// fieldbus master, which lives in Tether's io plane — they are a
// documented gap.  The *general* IOF blocks are meaningful and
// are implemented here over the package variable table:
//   IOF_GetBoxCount / IOF_GetBoxNameByAddr / IOF_GetBoxAddrByName /
//   IOF_GetDeviceCount / IOF_GetDeviceName.
// Documented differences:
//   - A "box" is an AT-bound variable (%I/%Q/%M) of the local
//     program, addressed by its image byte (and bit for BOOLs).
//     There is one local device (the PLC) — no fieldbus devices.
//   - IOF_DeviceReset and the *Ex/NetId/DeviceID variants need the
//     I/O server: they report a documented unsupported error
//     instead of pretending to reset hardware.

FUNCTION_BLOCK IOF_GetBoxCount
VAR_INPUT
    bExecute : BOOL;
    sNetId : STRING[23];
END_VAR
VAR_OUTPUT
    nCount : UDINT;
    bBusy : BOOL;
    bDone : BOOL;
    bError : BOOL;
    nErrId : UDINT;
END_VAR
VAR
    iof : FB_Iof;
    prev : BOOL;
END_VAR
    bBusy := FALSE; bDone := FALSE; bError := FALSE; nErrId := 0;
    IF bExecute AND NOT prev THEN
        bBusy := TRUE;
        iof.OP := 1;
        iof();
        bBusy := FALSE;
        IF iof.STATUS = 0 THEN
            bDone := TRUE; nCount := iof.COUNT;
        ELSE
            bError := TRUE; nErrId := iof.ERRID;
        END_IF;
    END_IF;
    prev := bExecute;
END_FUNCTION_BLOCK

FUNCTION_BLOCK IOF_GetBoxNameByAddr
VAR_INPUT
    bExecute : BOOL;
    sNetId : STRING[23];
    nRegion : UDINT;            // 0=%I 1=%Q 2=%M
    nAddr : UDINT;              // image byte
END_VAR
VAR_OUTPUT
    sName : STRING[63];
    bBusy : BOOL;
    bDone : BOOL;
    bError : BOOL;
    nErrId : UDINT;
END_VAR
VAR
    iof : FB_Iof;
    prev : BOOL;
    i : UDINT;
    n : UDINT;
    found : BOOL;
END_VAR
    bBusy := FALSE; bDone := FALSE; bError := FALSE; nErrId := 0;
    IF bExecute AND NOT prev THEN
        bBusy := TRUE;
        // scan the box list for the requested (region, addr)
        iof.OP := 1;
        iof();
        n := iof.COUNT;
        found := FALSE;
        i := 0;
        WHILE i < n AND NOT found DO
            iof.OP := 2; iof.IDX := i;
            iof();
            IF iof.FOUND AND iof.REGION = nRegion AND iof.ADDR = nAddr THEN
                sName := iof.NAME;
                found := TRUE;
            END_IF;
            i := i + 1;
        END_WHILE;
        bBusy := FALSE;
        IF found THEN
            bDone := TRUE;
        ELSE
            bError := TRUE; nErrId := 2;
        END_IF;
    END_IF;
    prev := bExecute;
END_FUNCTION_BLOCK

FUNCTION_BLOCK IOF_GetBoxAddrByName
VAR_INPUT
    bExecute : BOOL;
    sNetId : STRING[23];
    sName : STRING[63];
END_VAR
VAR_OUTPUT
    nRegion : UDINT;
    nAddr : UDINT;
    nUnit : UDINT;
    bBusy : BOOL;
    bDone : BOOL;
    bError : BOOL;
    nErrId : UDINT;
END_VAR
VAR
    iof : FB_Iof;
    prev : BOOL;
END_VAR
    bBusy := FALSE; bDone := FALSE; bError := FALSE; nErrId := 0;
    IF bExecute AND NOT prev THEN
        bBusy := TRUE;
        iof.OP := 3; iof.NAME := sName;
        iof();
        bBusy := FALSE;
        IF iof.STATUS = 0 AND iof.FOUND THEN
            bDone := TRUE;
            nRegion := iof.REGION;
            nAddr := iof.ADDR;
            nUnit := iof.UNIT;
        ELSE
            bError := TRUE; nErrId := iof.ERRID;
        END_IF;
    END_IF;
    prev := bExecute;
END_FUNCTION_BLOCK

FUNCTION_BLOCK IOF_GetDeviceCount
VAR_INPUT
    bExecute : BOOL;
    sNetId : STRING[23];
END_VAR
VAR_OUTPUT
    nCount : UDINT;
    bBusy : BOOL;
    bDone : BOOL;
    bError : BOOL;
    nErrId : UDINT;
END_VAR
VAR
    iof : FB_Iof;
    prev : BOOL;
END_VAR
    bBusy := FALSE; bDone := FALSE; bError := FALSE; nErrId := 0;
    IF bExecute AND NOT prev THEN
        bBusy := TRUE;
        iof.OP := 4;
        iof();
        bBusy := FALSE;
        IF iof.STATUS = 0 THEN
            bDone := TRUE; nCount := iof.COUNT;
        ELSE
            bError := TRUE; nErrId := iof.ERRID;
        END_IF;
    END_IF;
    prev := bExecute;
END_FUNCTION_BLOCK

FUNCTION_BLOCK IOF_GetDeviceName
VAR_INPUT
    bExecute : BOOL;
    sNetId : STRING[23];
    nDevId : UDINT;
END_VAR
VAR_OUTPUT
    sName : STRING[63];
    bBusy : BOOL;
    bDone : BOOL;
    bError : BOOL;
    nErrId : UDINT;
END_VAR
VAR
    iof : FB_Iof;
    prev : BOOL;
END_VAR
    bBusy := FALSE; bDone := FALSE; bError := FALSE; nErrId := 0;
    IF bExecute AND NOT prev THEN
        bBusy := TRUE;
        iof.OP := 5;
        iof();
        bBusy := FALSE;
        IF iof.STATUS = 0 AND nDevId = 0 THEN
            bDone := TRUE; sName := iof.VAL;
        ELSE
            bError := TRUE; nErrId := 3;
        END_IF;
    END_IF;
    prev := bExecute;
END_FUNCTION_BLOCK

// ---- host-domain operations: documented unsupported ----
FUNCTION_BLOCK IOF_DeviceReset
VAR_INPUT
    bExecute : BOOL;
    sNetId : STRING[23];
    nDevId : UDINT;
END_VAR
VAR_OUTPUT
    bBusy : BOOL;
    bDone : BOOL;
    bError : BOOL;
    nErrId : UDINT;
END_VAR
VAR
    prev : BOOL;
END_VAR
    bBusy := FALSE; bDone := FALSE; bError := FALSE; nErrId := 0;
    IF bExecute AND NOT prev THEN
        // resets are performed by the I/O plane (Tether), not the PLC
        bError := TRUE; nErrId := 16#8001;
    END_IF;
    prev := bExecute;
END_FUNCTION_BLOCK

FUNCTION_BLOCK IOF_GetBoxAddrByNameEx
VAR_INPUT
    bExecute : BOOL;
    sNetId : STRING[23];
    sName : STRING[63];
END_VAR
VAR_OUTPUT
    nRegion : UDINT;
    nAddr : UDINT;
    nUnit : UDINT;
    nBoxType : UDINT;
    bBusy : BOOL;
    bDone : BOOL;
    bError : BOOL;
    nErrId : UDINT;
END_VAR
VAR
    byName : IOF_GetBoxAddrByName;
END_VAR
    byName.bExecute := bExecute;
    byName.sNetId := sNetId;
    byName.sName := sName;
    byName();
    nRegion := byName.nRegion;
    nAddr := byName.nAddr;
    nUnit := byName.nUnit;
    nBoxType := 0;              // no terminal-type model in the PLC
    bBusy := byName.bBusy;
    bDone := byName.bDone;
    bError := byName.bError;
    nErrId := byName.nErrId;
END_FUNCTION_BLOCK

FUNCTION_BLOCK IOF_GetBoxNetId
VAR_INPUT
    bExecute : BOOL;
    nRegion : UDINT;
    nAddr : UDINT;
END_VAR
VAR_OUTPUT
    sNetId : STRING[23];
    bBusy : BOOL;
    bDone : BOOL;
    bError : BOOL;
    nErrId : UDINT;
END_VAR
VAR
    prev : BOOL;
END_VAR
    bBusy := FALSE; bDone := FALSE; bError := FALSE; nErrId := 0;
    IF bExecute AND NOT prev THEN
        sNetId := '127.0.0.1.1.1';   // the local PLC is the only device
        bDone := TRUE;
    END_IF;
    prev := bExecute;
END_FUNCTION_BLOCK

FUNCTION_BLOCK IOF_GetDeviceNetId
VAR_INPUT
    bExecute : BOOL;
    nDevId : UDINT;
END_VAR
VAR_OUTPUT
    sNetId : STRING[23];
    bBusy : BOOL;
    bDone : BOOL;
    bError : BOOL;
    nErrId : UDINT;
END_VAR
VAR
    prev : BOOL;
END_VAR
    bBusy := FALSE; bDone := FALSE; bError := FALSE; nErrId := 0;
    IF bExecute AND NOT prev THEN
        sNetId := '127.0.0.1.1.1';
        bDone := TRUE;
    END_IF;
    prev := bExecute;
END_FUNCTION_BLOCK

FUNCTION_BLOCK IOF_GetDeviceIDByName
VAR_INPUT
    bExecute : BOOL;
    sNetId : STRING[23];
    sName : STRING[63];
END_VAR
VAR_OUTPUT
    nDevId : UDINT;
    bBusy : BOOL;
    bDone : BOOL;
    bError : BOOL;
    nErrId : UDINT;
END_VAR
VAR
    prev : BOOL;
END_VAR
    bBusy := FALSE; bDone := FALSE; bError := FALSE; nErrId := 0;
    IF bExecute AND NOT prev THEN
        // single local device, id 0
        nDevId := 0;
        bDone := TRUE;
    END_IF;
    prev := bExecute;
END_FUNCTION_BLOCK

FUNCTION_BLOCK IOF_GetDeviceIDs
VAR_INPUT
    bExecute : BOOL;
    sNetId : STRING[23];
END_VAR
VAR_OUTPUT
    nDevId : UDINT;
    nCount : UDINT;
    bBusy : BOOL;
    bDone : BOOL;
    bError : BOOL;
    nErrId : UDINT;
END_VAR
VAR
    prev : BOOL;
END_VAR
    bBusy := FALSE; bDone := FALSE; bError := FALSE; nErrId := 0;
    IF bExecute AND NOT prev THEN
        nDevId := 0; nCount := 1;
        bDone := TRUE;
    END_IF;
    prev := bExecute;
END_FUNCTION_BLOCK

FUNCTION_BLOCK IOF_GetDeviceInfoByName
VAR_INPUT
    bExecute : BOOL;
    sNetId : STRING[23];
    sName : STRING[63];
END_VAR
VAR_OUTPUT
    nDevId : UDINT;
    nDevType : UDINT;
    bBusy : BOOL;
    bDone : BOOL;
    bError : BOOL;
    nErrId : UDINT;
END_VAR
VAR
    prev : BOOL;
END_VAR
    bBusy := FALSE; bDone := FALSE; bError := FALSE; nErrId := 0;
    IF bExecute AND NOT prev THEN
        nDevId := 0; nDevType := 0;
        bDone := TRUE;
    END_IF;
    prev := bExecute;
END_FUNCTION_BLOCK

(* ---- tc2_mbus.st ---- *)
// tc2_mbus.st — wired M-Bus (EN 13757) metering-master surface
// (TwinCAT Tc3_MBus/TF6681-ish shape) over the tplc-mbus service +
// FB_Mbus builtin.
//
// The PLC is the M-Bus master over an opt-in serial port (2400 8E1):
// FB_MbusOpen opens the UART; FB_MbusShort carries the short frames
// (SND_NKE 0x40, REQ_UD2 0x5B, REQ_UD1 0x7B); FB_MbusLong carries
// long frames (SND_UD etc.); FB_MbusReceive polls for a response
// (E5 ack or a 68.. long frame); FB_MbusStatus reports counters.
//
// Payload fields are raw bytes bounded STRING[255] — the caller
// composes/parses the M-Bus DIF/VIF record.  Secondary addressing,
// the application-layer record decode, and the collision/FDB
// handling a full master does are honest gaps for a later tranche.

// ---- FB_MbusOpen: open the serial port (2400 8E1) ----
FUNCTION_BLOCK FB_MbusOpen
VAR_INPUT
    Execute : BOOL;
    Path : STRING[127];
END_VAR
VAR_OUTPUT
    Done : BOOL;
    Error : BOOL;
    ErrorID : UDINT;
    PortHdl : UDINT;
END_VAR
VAR
    ch : FB_Mbus;
    exPrev : BOOL;
END_VAR
    Done := FALSE;
    Error := FALSE;
    ErrorID := 0;
    IF Execute AND NOT exPrev THEN
        ch.OP := 1;
        ch.PATH := Path;
        ch();
        IF ch.STATUS = 0 THEN
            Done := TRUE;
            PortHdl := ch.HANDLE;
        ELSE
            Error := TRUE;
            ErrorID := ch.ERRID;
        END_IF;
    END_IF;
    exPrev := Execute;
END_FUNCTION_BLOCK

// ---- FB_MbusClose: release the serial port ----
FUNCTION_BLOCK FB_MbusClose
VAR_INPUT
    Execute : BOOL;
    PortHdl : UDINT;
END_VAR
VAR_OUTPUT
    Done : BOOL;
    Error : BOOL;
    ErrorID : UDINT;
END_VAR
VAR
    ch : FB_Mbus;
    exPrev : BOOL;
END_VAR
    Done := FALSE;
    Error := FALSE;
    ErrorID := 0;
    IF Execute AND NOT exPrev THEN
        ch.OP := 2;
        ch.HANDLE := PortHdl;
        ch();
        IF ch.STATUS = 0 THEN
            Done := TRUE;
        ELSE
            Error := TRUE;
            ErrorID := ch.ERRID;
        END_IF;
    END_IF;
    exPrev := Execute;
END_FUNCTION_BLOCK

// ---- FB_MbusShort: short frame (SND_NKE/REQ_UD2/REQ_UD1) ----
FUNCTION_BLOCK FB_MbusShort
VAR_INPUT
    Execute : BOOL;
    PortHdl : UDINT;
    Control : UDINT;
    Address : UDINT;
END_VAR
VAR_OUTPUT
    Done : BOOL;
    Error : BOOL;
    ErrorID : UDINT;
END_VAR
VAR
    ch : FB_Mbus;
    exPrev : BOOL;
END_VAR
    Done := FALSE;
    Error := FALSE;
    ErrorID := 0;
    IF Execute AND NOT exPrev THEN
        ch.OP := 4;
        ch.HANDLE := PortHdl;
        ch.CONTROL := Control;
        ch.ADDRESS := Address;
        ch();
        IF ch.STATUS = 0 THEN
            Done := TRUE;
        ELSE
            Error := TRUE;
            ErrorID := ch.ERRID;
        END_IF;
    END_IF;
    exPrev := Execute;
END_FUNCTION_BLOCK

// ---- FB_MbusLong: long frame (SND_UD etc.) ----
FUNCTION_BLOCK FB_MbusLong
VAR_INPUT
    Execute : BOOL;
    PortHdl : UDINT;
    Control : UDINT;
    Address : UDINT;
    Ci : UDINT;
    Data : STRING[255];
END_VAR
VAR_OUTPUT
    Done : BOOL;
    Error : BOOL;
    ErrorID : UDINT;
END_VAR
VAR
    ch : FB_Mbus;
    exPrev : BOOL;
END_VAR
    Done := FALSE;
    Error := FALSE;
    ErrorID := 0;
    IF Execute AND NOT exPrev THEN
        ch.OP := 5;
        ch.HANDLE := PortHdl;
        ch.CONTROL := Control;
        ch.ADDRESS := Address;
        ch.CI := Ci;
        ch.DATA := Data;
        ch();
        IF ch.STATUS = 0 THEN
            Done := TRUE;
        ELSE
            Error := TRUE;
            ErrorID := ch.ERRID;
        END_IF;
    END_IF;
    exPrev := Execute;
END_FUNCTION_BLOCK

// ---- FB_MbusReceive: poll for a response (E5 / 68..) ----
FUNCTION_BLOCK FB_MbusReceive
VAR_INPUT
    Execute : BOOL;
    PortHdl : UDINT;
END_VAR
VAR_OUTPUT
    Done : BOOL;
    Message : BOOL;
    Error : BOOL;
    ErrorID : UDINT;
    Kind : UDINT;
    Payload : STRING[255];
END_VAR
VAR
    ch : FB_Mbus;
END_VAR
    Done := FALSE;
    Message := FALSE;
    Error := FALSE;
    ErrorID := 0;
    IF Execute THEN
        ch.OP := 6;
        ch.HANDLE := PortHdl;
        ch();
        IF ch.STATUS = 1 THEN
            Done := TRUE;               // NOMSG: still waiting
        ELSIF ch.STATUS >= 0 THEN
            Done := TRUE;
            Message := TRUE;
            Kind := ch.KIND;
            Payload := ch.RXPAYLOAD;
        ELSE
            Error := TRUE;
            ErrorID := ch.ERRID;
        END_IF;
    END_IF;
END_FUNCTION_BLOCK

// ---- FB_MbusStatus: frame counters + state ----
FUNCTION_BLOCK FB_MbusStatus
VAR_INPUT
    Execute : BOOL;
    PortHdl : UDINT;
END_VAR
VAR_OUTPUT
    Done : BOOL;
    Error : BOOL;
    ErrorID : UDINT;
    State : DINT;
    TxTotal : UDINT;
    RxTotal : UDINT;
    LastErr : DINT;
END_VAR
VAR
    ch : FB_Mbus;
END_VAR
    Done := FALSE;
    Error := FALSE;
    ErrorID := 0;
    IF Execute THEN
        ch.OP := 3;
        ch.HANDLE := PortHdl;
        ch();
        IF ch.STATUS = 0 THEN
            Done := TRUE;
            State := ch.STATE;
            TxTotal := ch.TXTOT;
            RxTotal := ch.RXTOT;
            LastErr := ch.LASTERR;
        ELSE
            Error := TRUE;
            ErrorID := ch.ERRID;
        END_IF;
    END_IF;
END_FUNCTION_BLOCK

(* ---- tc2_mc2.st ---- *)
// Tc2_MC2 — TwinCAT PLCopen motion function blocks over the
// builtin FB_MotionAxis (tplc-motion service), a simulated
// CiA402/DS402-shaped axis pool.
//
// AXIS_REF mapping: TwinCAT's AXIS_REF is a large structure
// (PlcToDrive/DriveToPlc sub-records, axis id, parameters). The
// simulated backend identifies an axis by a bounded UDINT handle
// returned from FB_MotionAxis OP=1 create, so the compat surface
// takes that handle as the `Axis` input. Position/velocity values
// are the backend's native int32 user units (TwinCAT uses LREAL
// engineering units; the LREAL<->int conversion is a documented
// gap). This file implements the axis-management blocks
// (MC_Power/MC_Reset/MC_SetPosition/MC_Read*), the point-to-point /
// velocity / stop / halt / homing / jog command blocks, and the
// modulo / override / axis-parameter FBs. The motion-command FBs
// drive the DS402 controlword command pattern (NewSetPoint for
// PP/HM, QuickStop for MC_Stop) and the mode/target objects;
// per-command Velocity/Acceleration/Deceleration inputs are
// accepted for signature compatibility but the simulated axis
// applies its configured dynamics limits.
// SPDX-License-Identifier: Apache-2.0 OR MPL-2.0

// DS402 object indices used by the wrappers.
// (declared as constants via VAR in each FB that needs them)

// ---- MC_Power: software enable of the axis ----
// Enable=TRUE drives the controlword to EnableOperation (0x000F);
// Enable=FALSE drives DisableVoltage (0x0000). The controlword is
// written only on an Enable transition (edge-triggered) so the
// motion-command FBs can layer NewSetPoint/QuickStop command bits
// on top without being overwritten every scan; the drive holds the
// commanded state. Status is TRUE once the axis reports CiA402
// OperationEnabled (state 0x27 = 39). Enable_Positive/
// Enable_Negative are accepted for signature compatibility; the
// simulated axis is bidirectional so only Enable gates power.
FUNCTION_BLOCK MC_Power
VAR_INPUT
    Enable : BOOL;
    Enable_Positive : BOOL;
    Enable_Negative : BOOL;
    Axis : UDINT;
END_VAR
VAR_OUTPUT
    Status : BOOL;
    Busy : BOOL;
    Error : BOOL;
    ErrorID : UDINT;
END_VAR
VAR
    ax : FB_MotionAxis;
    enPrev : BOOL;
END_VAR
    // advance dynamics once per scan
    ax.OP := 3; ax();
    ax.AXIS := Axis;
    // edge-trigger the enable command so command FBs own the
    // controlword's command bits between transitions
    IF Enable <> enPrev THEN
        ax.OP := 5;
        ax.INDEX := 16#6040;
        IF Enable THEN
            ax.VALUE := 16#000F;
        ELSE
            ax.VALUE := 0;
        END_IF;
        ax();
        enPrev := Enable;
    END_IF;
    // snapshot for Status (CiA402 state in STATUS for OP=6)
    ax.OP := 6;
    ax();
    Status := (ax.STATUS = 39);
    Busy := FALSE;
    Error := FALSE;
    ErrorID := 0;
END_FUNCTION_BLOCK

// ---- MC_Reset: reset the axis (fault reset controlword bit) ----
// Execute rising edge pulses controlword bit7 (FaultReset,
// 0x0080) onto the enable command for one scan, then releases it
// the next scan. To avoid fighting MC_Power over 0x6040, the
// controlword is only written during that two-scan window; on
// other scans the FB leaves the controlword to MC_Power. Done
// reports the reset write succeeded.
FUNCTION_BLOCK MC_Reset
VAR_INPUT
    Execute : BOOL;
    Axis : UDINT;
END_VAR
VAR_OUTPUT
    Done : BOOL;
    Busy : BOOL;
    Error : BOOL;
    ErrorID : UDINT;
END_VAR
VAR
    ax : FB_MotionAxis;
    edge : BOOL;
    rst : BOOL;
    rel : BOOL;
END_VAR
    edge := Execute AND NOT rst;
    rst := Execute;
    ax.AXIS := Axis;
    ax.OP := 3; ax();   // advance dynamics/state
    IF edge OR rel THEN
        ax.OP := 5;
        ax.INDEX := 16#6040;
        IF edge THEN
            ax.VALUE := 16#008F;   // FaultReset | EnableOperation
        ELSE
            ax.VALUE := 16#000F;   // release reset, stay enabled
        END_IF;
        ax();
        rel := edge;              // next scan releases bit7
        Done := (edge AND ax.STATUS = 0);
    ELSE
        rel := FALSE;
        Done := FALSE;
    END_IF;
    Busy := FALSE;
    Error := FALSE;
    ErrorID := 0;
END_FUNCTION_BLOCK

// ---- MC_SetPosition: preset the axis position ----
// Execute rising edge writes PositionActualValue (0x6064): the
// absolute value, or current+Position when Mode=TRUE (relative).
// Position is int32 user units (LREAL engineering units is a gap).
FUNCTION_BLOCK MC_SetPosition
VAR_INPUT
    Execute : BOOL;
    Position : DINT;
    Mode : BOOL;
    Axis : UDINT;
END_VAR
VAR_OUTPUT
    Done : BOOL;
    Busy : BOOL;
    Error : BOOL;
    ErrorID : UDINT;
END_VAR
VAR
    ax : FB_MotionAxis;
    edge : BOOL;
    rst : BOOL;
    cur : DINT;
    np : DINT;
END_VAR
    edge := Execute AND NOT rst;
    rst := Execute;
    // Position write is edge-triggered only; rewriting every scan would
    // re-apply a stale Position input and revert later moves.
    IF edge THEN
        np := Position;
        IF Mode THEN
            // relative: read current actual position first
            ax.AXIS := Axis;
            ax.OP := 4;
            ax.INDEX := 16#6064;
            ax();
            cur := ax.VALUE;
            np := cur + Position;
        END_IF;
        ax.AXIS := Axis;
        ax.OP := 5;
        ax.INDEX := 16#6064;
        ax.VALUE := np;
        ax();
        IF ax.STATUS = 0 THEN
            Done := TRUE;
        ELSE
            Done := FALSE;
            Error := TRUE;
            ErrorID := ax.STATUS;
        END_IF;
    ELSE
        Done := FALSE;
        Error := FALSE;
        ErrorID := 0;
    END_IF;
    Busy := FALSE;
END_FUNCTION_BLOCK

// ---- MC_ReadActualPosition: read position actual value ----
// Enable=TRUE reads cyclically; Valid/Position carry the value.
FUNCTION_BLOCK MC_ReadActualPosition
VAR_INPUT
    Enable : BOOL;
    Axis : UDINT;
END_VAR
VAR_OUTPUT
    Valid : BOOL;
    Position : DINT;
    Busy : BOOL;
END_VAR
VAR
    ax : FB_MotionAxis;
END_VAR
    ax.OP := 3; ax();
    ax.AXIS := Axis;
    ax.OP := 4;
    ax.INDEX := 16#6064;
    ax();
    IF Enable AND ax.STATUS = 0 THEN
        Valid := TRUE;
        Position := ax.VALUE;
    ELSE
        Valid := FALSE;
        Position := 0;
    END_IF;
    Busy := FALSE;
END_FUNCTION_BLOCK

// ---- MC_ReadActualVelocity: read velocity actual value ----
FUNCTION_BLOCK MC_ReadActualVelocity
VAR_INPUT
    Enable : BOOL;
    Axis : UDINT;
END_VAR
VAR_OUTPUT
    Valid : BOOL;
    Velocity : DINT;
    Busy : BOOL;
END_VAR
VAR
    ax : FB_MotionAxis;
END_VAR
    ax.OP := 3; ax();
    ax.AXIS := Axis;
    ax.OP := 4;
    ax.INDEX := 16#606C;
    ax();
    IF Enable AND ax.STATUS = 0 THEN
        Valid := TRUE;
        Velocity := ax.VALUE;
    ELSE
        Valid := FALSE;
        Velocity := 0;
    END_IF;
    Busy := FALSE;
END_FUNCTION_BLOCK

// ---- MC_ReadAxisError: read the axis error code ----
// Valid=TRUE when the read succeeded; AxisErrorID is the DS402
// error code object (0x603F), 0 when no fault is latched.
FUNCTION_BLOCK MC_ReadAxisError
VAR_INPUT
    Enable : BOOL;
    Axis : UDINT;
END_VAR
VAR_OUTPUT
    Valid : BOOL;
    AxisErrorID : DINT;
    Busy : BOOL;
END_VAR
VAR
    ax : FB_MotionAxis;
END_VAR
    ax.OP := 3; ax();
    ax.AXIS := Axis;
    ax.OP := 4;
    ax.INDEX := 16#603F;
    ax();
    IF Enable AND ax.STATUS = 0 THEN
        Valid := TRUE;
        AxisErrorID := ax.VALUE;
    ELSE
        Valid := FALSE;
        AxisErrorID := 0;
    END_IF;
    Busy := FALSE;
END_FUNCTION_BLOCK

// ---- MC_ReadStatus: read the axis operating state ----
// Reports the PLCopen operating state derived from the CiA402
// status, mode display, actual velocity and fault flags:
//   0=Disabled, 1=Standstill, 2=Homing, 3=DiscreteMotion,
//   4=ContinuousMotion, 6=Stopping, 7=ErrorStop (-1=read fail).
// (5=SynchronizedMotion is reserved for gearing/camming, not yet
// produced.) Valid signals a successful read.
FUNCTION_BLOCK MC_ReadStatus
VAR_INPUT
    Enable : BOOL;
    Axis : UDINT;
END_VAR
VAR_OUTPUT
    Valid : BOOL;
    OperatingState : INT;
    Busy : BOOL;
END_VAR
VAR
    ax : FB_MotionAxis;
    stt : DINT;
    md : DINT;
    tr : DINT;
    va : DINT;
END_VAR
    ax.OP := 3; ax();
    ax.AXIS := Axis;
    ax.OP := 6;
    ax();
    IF Enable AND ax.STATUS >= 0 THEN
        Valid := TRUE;
        stt := ax.STATUS;            // CiA402 state
        md := ax.MODE;               // mode of operation display
        tr := ax.TARGET_REACHED;
        va := ax.VEL_ACTUAL;
        IF ax.FAULT <> 0 OR stt = 8 OR stt = 15 THEN
            OperatingState := 7;     // ErrorStop (fault latched)
        ELSIF stt = 7 THEN
            OperatingState := 6;     // Stopping (QuickStopActive)
        ELSIF stt <> 39 THEN
            OperatingState := 0;     // Disabled / not ready
        ELSIF md = 6 THEN
            OperatingState := 2;     // Homing
        ELSIF md = 1 AND tr = 0 THEN
            OperatingState := 3;     // DiscreteMotion (PP move active)
        ELSIF (md = 2 OR md = 3 OR md = 8 OR md = 9 OR md = 10)
              AND va <> 0 THEN
            OperatingState := 4;     // ContinuousMotion (moving)
        ELSE
            OperatingState := 1;     // Standstill (enabled, at rest)
        END_IF;
    ELSE
        Valid := FALSE;
        OperatingState := -1;
    END_IF;
    Busy := FALSE;
END_FUNCTION_BLOCK

// ================================================================== //
// Motion-command FBs. Each drives the DS402 controlword command
// pattern on its Execute edge: PP/HM modes pulse NewSetPoint
// (0x0010) with the enable pattern for one scan then release to
// 0x000F; velocity modes write mode+target velocity under the
// enable pattern; MC_Stop commands QuickStop (controlword QS bit
// cleared); MC_Halt ramps profile-velocity to zero. The controlword
// is written only on the command edge (plus the single NSP release
// scan), so MC_Power's edge-triggered enable is not fought and a
// later MC_Stop/MC_Power transition can override a running command.
// ================================================================== //

// ---- MC_MoveAbsolute: absolute point-to-point move (PP mode) ----
// Execute edge: mode=ProfilePosition, TargetPosition=Position,
// controlword=EnableOperation|NewSetPoint (0x001F). Done when the
// axis reports TargetReached (statusword bit 0x0400). Velocity/
// Acceleration/Deceleration are signature-compatible; the axis
// applies its configured dynamics.
FUNCTION_BLOCK MC_MoveAbsolute
VAR_INPUT
    Execute : BOOL;
    Position : DINT;
    Velocity : DINT;
    Acceleration : DINT;
    Deceleration : DINT;
    Axis : UDINT;
END_VAR
VAR_OUTPUT
    Done : BOOL;
    Busy : BOOL;
    CommandAborted : BOOL;
    Error : BOOL;
    ErrorID : UDINT;
END_VAR
VAR
    ax : FB_MotionAxis;
    exPrev : BOOL;
    exEdge : BOOL;
    active : BOOL;
    rel : BOOL;
END_VAR
    ax.AXIS := Axis;
    ax.OP := 3; ax();
    exEdge := Execute AND NOT exPrev; exPrev := Execute;
    Done := FALSE; CommandAborted := FALSE; Error := FALSE; ErrorID := 0;
    IF NOT active AND exEdge THEN
        ax.OP := 5; ax.INDEX := 16#6060; ax.VALUE := 1; ax();
        ax.OP := 5; ax.INDEX := 16#607A; ax.VALUE := Position; ax();
        ax.OP := 5; ax.INDEX := 16#6040; ax.VALUE := 16#001F; ax();
        IF ax.STATUS = 0 THEN
            active := TRUE; rel := TRUE;
        ELSE
            Error := TRUE; ErrorID := ax.ERRID;
        END_IF;
    ELSIF active THEN
        IF rel THEN
            ax.OP := 5; ax.INDEX := 16#6040; ax.VALUE := 16#000F; ax();
            rel := FALSE;
        END_IF;
        ax.OP := 6; ax();
        IF ax.STATUS < 0 THEN
            Error := TRUE; ErrorID := ax.ERRID; active := FALSE;
        ELSIF ax.TARGET_REACHED = 1 THEN
            Done := TRUE; active := FALSE;
        END_IF;
    END_IF
    Busy := active;
END_FUNCTION_BLOCK

// ---- MC_MoveRelative: relative point-to-point move (PP mode) ----
// Execute edge reads PositionActualValue, adds Distance, then runs
// the same PP/NewSetPoint sequence as MC_MoveAbsolute.
FUNCTION_BLOCK MC_MoveRelative
VAR_INPUT
    Execute : BOOL;
    Distance : DINT;
    Velocity : DINT;
    Acceleration : DINT;
    Deceleration : DINT;
    Axis : UDINT;
END_VAR
VAR_OUTPUT
    Done : BOOL;
    Busy : BOOL;
    CommandAborted : BOOL;
    Error : BOOL;
    ErrorID : UDINT;
END_VAR
VAR
    ax : FB_MotionAxis;
    exPrev : BOOL;
    exEdge : BOOL;
    active : BOOL;
    rel : BOOL;
    cur : DINT;
END_VAR
    ax.AXIS := Axis;
    ax.OP := 3; ax();
    exEdge := Execute AND NOT exPrev; exPrev := Execute;
    Done := FALSE; CommandAborted := FALSE; Error := FALSE; ErrorID := 0;
    IF NOT active AND exEdge THEN
        ax.OP := 4; ax.INDEX := 16#6064; ax();   // read pos actual
        cur := ax.VALUE;
        ax.OP := 5; ax.INDEX := 16#6060; ax.VALUE := 1; ax();
        ax.OP := 5; ax.INDEX := 16#607A; ax.VALUE := cur + Distance; ax();
        ax.OP := 5; ax.INDEX := 16#6040; ax.VALUE := 16#001F; ax();
        IF ax.STATUS = 0 THEN
            active := TRUE; rel := TRUE;
        ELSE
            Error := TRUE; ErrorID := ax.ERRID;
        END_IF;
    ELSIF active THEN
        IF rel THEN
            ax.OP := 5; ax.INDEX := 16#6040; ax.VALUE := 16#000F; ax();
            rel := FALSE;
        END_IF;
        ax.OP := 6; ax();
        IF ax.STATUS < 0 THEN
            Error := TRUE; ErrorID := ax.ERRID; active := FALSE;
        ELSIF ax.TARGET_REACHED = 1 THEN
            Done := TRUE; active := FALSE;
        END_IF;
    END_IF
    Busy := active;
END_FUNCTION_BLOCK

// ---- MC_MoveVelocity: endless travel at Velocity (PV mode) ----
// Execute edge: mode=ProfileVelocity, TargetVelocity=Velocity,
// controlword=EnableOperation. The axis ramps to the target velocity
// and holds it; the move ends via MC_Stop/MC_Halt. ContinuousUpdate
// rewrites TargetVelocity each scan for live dynamics changes.
// InVelocity reports TargetReached (|vel-target| within window).
FUNCTION_BLOCK MC_MoveVelocity
VAR_INPUT
    Execute : BOOL;
    ContinuousUpdate : BOOL;
    Velocity : DINT;
    Acceleration : DINT;
    Deceleration : DINT;
    Axis : UDINT;
END_VAR
VAR_OUTPUT
    InVelocity : BOOL;
    Busy : BOOL;
    CommandAborted : BOOL;
    Error : BOOL;
    ErrorID : UDINT;
END_VAR
VAR
    ax : FB_MotionAxis;
    exPrev : BOOL;
    exEdge : BOOL;
    engaged : BOOL;
END_VAR
    ax.AXIS := Axis;
    ax.OP := 3; ax();
    exEdge := Execute AND NOT exPrev; exPrev := Execute;
    InVelocity := FALSE; CommandAborted := FALSE; Error := FALSE; ErrorID := 0;
    IF exEdge THEN
        ax.OP := 5; ax.INDEX := 16#6040; ax.VALUE := 16#000F; ax();
        ax.OP := 5; ax.INDEX := 16#6060; ax.VALUE := 3; ax();
        ax.OP := 5; ax.INDEX := 16#60FF; ax.VALUE := Velocity; ax();
        engaged := TRUE;
    END_IF
    IF engaged AND ContinuousUpdate THEN
        ax.OP := 5; ax.INDEX := 16#60FF; ax.VALUE := Velocity; ax();
    END_IF
    IF engaged THEN
        ax.OP := 6; ax();
        IF ax.STATUS < 0 THEN
            Error := TRUE; ErrorID := ax.ERRID; engaged := FALSE;
        ELSE
            InVelocity := (ax.TARGET_REACHED = 1);
        END_IF
    END_IF
    Busy := engaged;
END_FUNCTION_BLOCK

// ---- MC_Stop: quick stop, locks the axis ----
// Execute edge commands QuickStop by clearing the controlword QS
// bit (write 0x000B = enable pattern without QuickStop-request).
// The drive decelerates to rest and holds QuickStopActive; Done
// reports when VelocityActualValue reaches zero. A later motion
// command re-asserts the enable pattern and resumes.
FUNCTION_BLOCK MC_Stop
VAR_INPUT
    Execute : BOOL;
    Deceleration : DINT;
    Axis : UDINT;
END_VAR
VAR_OUTPUT
    Done : BOOL;
    Busy : BOOL;
    CommandAborted : BOOL;
    Error : BOOL;
    ErrorID : UDINT;
END_VAR
VAR
    ax : FB_MotionAxis;
    exPrev : BOOL;
    exEdge : BOOL;
    active : BOOL;
END_VAR
    ax.AXIS := Axis;
    ax.OP := 3; ax();
    exEdge := Execute AND NOT exPrev; exPrev := Execute;
    Done := FALSE; CommandAborted := FALSE; Error := FALSE; ErrorID := 0;
    IF NOT active AND exEdge THEN
        ax.OP := 5; ax.INDEX := 16#6040; ax.VALUE := 16#000B; ax();
        IF ax.STATUS = 0 THEN
            active := TRUE;
        ELSE
            Error := TRUE; ErrorID := ax.ERRID;
        END_IF;
    ELSIF active THEN
        ax.OP := 6; ax();
        IF ax.STATUS < 0 THEN
            Error := TRUE; ErrorID := ax.ERRID; active := FALSE;
        ELSIF ax.VEL_ACTUAL = 0 THEN
            Done := TRUE; active := FALSE;
        END_IF;
    END_IF
    Busy := active;
END_FUNCTION_BLOCK

// ---- MC_Halt: controlled stop with ramp (stays enabled) ----
// Execute edge: mode=ProfileVelocity, TargetVelocity=0 under the
// enable pattern, so the axis ramps to rest at its configured
// deceleration and remains OperationEnabled. Done when velocity
// reaches zero. Unlike MC_Stop the axis is not locked and a new
// command can resume immediately.
FUNCTION_BLOCK MC_Halt
VAR_INPUT
    Execute : BOOL;
    Deceleration : DINT;
    Axis : UDINT;
END_VAR
VAR_OUTPUT
    Done : BOOL;
    Busy : BOOL;
    CommandAborted : BOOL;
    Error : BOOL;
    ErrorID : UDINT;
END_VAR
VAR
    ax : FB_MotionAxis;
    exPrev : BOOL;
    exEdge : BOOL;
    active : BOOL;
END_VAR
    ax.AXIS := Axis;
    ax.OP := 3; ax();
    exEdge := Execute AND NOT exPrev; exPrev := Execute;
    Done := FALSE; CommandAborted := FALSE; Error := FALSE; ErrorID := 0;
    IF NOT active AND exEdge THEN
        ax.OP := 5; ax.INDEX := 16#6040; ax.VALUE := 16#000F; ax();
        ax.OP := 5; ax.INDEX := 16#6060; ax.VALUE := 3; ax();
        ax.OP := 5; ax.INDEX := 16#60FF; ax.VALUE := 0; ax();
        active := TRUE;
    ELSIF active THEN
        ax.OP := 6; ax();
        IF ax.STATUS < 0 THEN
            Error := TRUE; ErrorID := ax.ERRID; active := FALSE;
        ELSIF ax.VEL_ACTUAL = 0 THEN
            Done := TRUE; active := FALSE;
        END_IF;
    END_IF
    Busy := active;
END_FUNCTION_BLOCK

// ---- MC_Home: homing move to the home offset (HM mode) ----
// Execute edge: writes HomeOffset=Position (0x607C, the reference
// position after homing), mode=Homing, controlword=enable|NewSet-
// Point. Done when the axis reports TargetReached/homing complete.
FUNCTION_BLOCK MC_Home
VAR_INPUT
    Execute : BOOL;
    Position : DINT;
    Velocity : DINT;
    Acceleration : DINT;
    Deceleration : DINT;
    Axis : UDINT;
END_VAR
VAR_OUTPUT
    Done : BOOL;
    Busy : BOOL;
    CommandAborted : BOOL;
    Error : BOOL;
    ErrorID : UDINT;
END_VAR
VAR
    ax : FB_MotionAxis;
    exPrev : BOOL;
    exEdge : BOOL;
    active : BOOL;
    rel : BOOL;
END_VAR
    ax.AXIS := Axis;
    ax.OP := 3; ax();
    exEdge := Execute AND NOT exPrev; exPrev := Execute;
    Done := FALSE; CommandAborted := FALSE; Error := FALSE; ErrorID := 0;
    IF NOT active AND exEdge THEN
        ax.OP := 5; ax.INDEX := 16#607C; ax.VALUE := Position; ax();
        ax.OP := 5; ax.INDEX := 16#6060; ax.VALUE := 6; ax();
        ax.OP := 5; ax.INDEX := 16#6040; ax.VALUE := 16#001F; ax();
        IF ax.STATUS = 0 THEN
            active := TRUE; rel := TRUE;
        ELSE
            Error := TRUE; ErrorID := ax.ERRID;
        END_IF;
    ELSIF active THEN
        IF rel THEN
            ax.OP := 5; ax.INDEX := 16#6040; ax.VALUE := 16#000F; ax();
            rel := FALSE;
        END_IF;
        ax.OP := 6; ax();
        IF ax.STATUS < 0 THEN
            Error := TRUE; ErrorID := ax.ERRID; active := FALSE;
        ELSIF ax.TARGET_REACHED = 1 THEN
            Done := TRUE; active := FALSE;
        END_IF;
    END_IF
    Busy := active;
END_FUNCTION_BLOCK

// ---- MC_Jog: manual jog while a direction key is held (PV mode) ----
// JogForward/JogBackwards are level inputs: while held the axis ramps
// to +/-Velocity in ProfileVelocity mode; on release TargetVelocity
// returns to 0 and the axis ramps to rest. Busy is TRUE while a key
// is held; Done pulses once the axis is back at rest after a jog.
// The mode is latched to ProfileVelocity on the first key press.
FUNCTION_BLOCK MC_Jog
VAR_INPUT
    JogForward : BOOL;
    JogBackwards : BOOL;
    Velocity : DINT;
    Axis : UDINT;
END_VAR
VAR_OUTPUT
    Done : BOOL;
    Busy : BOOL;
    Error : BOOL;
    ErrorID : UDINT;
END_VAR
VAR
    ax : FB_MotionAxis;
    modeSet : BOOL;
    wasMoving : BOOL;
    key : BOOL;
    stopped : BOOL;
END_VAR
    ax.AXIS := Axis;
    ax.OP := 3; ax();
    key := JogForward OR JogBackwards;
    Done := FALSE; Error := FALSE; ErrorID := 0;
    IF key AND NOT modeSet THEN
        ax.OP := 5; ax.INDEX := 16#6040; ax.VALUE := 16#000F; ax();
        ax.OP := 5; ax.INDEX := 16#6060; ax.VALUE := 3; ax();
        modeSet := TRUE;
    END_IF
    // velocity target follows the held key every scan
    IF JogForward THEN
        ax.OP := 5; ax.INDEX := 16#60FF; ax.VALUE := Velocity; ax();
    ELSIF JogBackwards THEN
        ax.OP := 5; ax.INDEX := 16#60FF; ax.VALUE := -Velocity; ax();
    ELSE
        ax.OP := 5; ax.INDEX := 16#60FF; ax.VALUE := 0; ax();
    END_IF
    ax.OP := 6; ax();
    stopped := (NOT key) AND (ax.VEL_ACTUAL = 0);
    IF stopped AND wasMoving THEN
        Done := TRUE;
    END_IF
    wasMoving := NOT stopped;
    Busy := NOT stopped;
END_FUNCTION_BLOCK

// ================================================================== //
// Tranche-4 blocks: modulo positioning, velocity override and the
// axis-parameter access FBs. The parameter FBs treat ParameterNumber
// as the DS402 object-dictionary index (0x0000..0xFFFF), giving
// generic object access through the PLCopen-style signature; the
// TwinCAT numeric parameter ids map onto indices in a real system,
// which is a documented simplification. Gearing/phasing/camming and
// hardware touch-probe latch need multi-axis coupling / latch
// objects the simulated backend does not expose — see README gaps.
// ================================================================== //

// ---- MC_MoveModulo: modulo positioning (PP mode) ----
// Position is the modulo target in [0,ModuloFactor). Direction
// selects the travel path: 0=shortest (default), 1=positive
// direction only, 2=negative direction only. The absolute target
// is computed from the current position so the axis lands on the
// requested modulo angle, then a standard PP/NewSetPoint move runs.
FUNCTION_BLOCK MC_MoveModulo
VAR_INPUT
    Execute : BOOL;
    Position : DINT;
    Velocity : DINT;
    Acceleration : DINT;
    Deceleration : DINT;
    Direction : INT;
    ModuloFactor : DINT;
    Axis : UDINT;
END_VAR
VAR_OUTPUT
    Done : BOOL;
    Busy : BOOL;
    CommandAborted : BOOL;
    Error : BOOL;
    ErrorID : UDINT;
END_VAR
VAR
    ax : FB_MotionAxis;
    exPrev : BOOL;
    exEdge : BOOL;
    active : BOOL;
    rel : BOOL;
    cur : DINT;
    tgt : DINT;
    delta : DINT;
    goal : DINT;
END_VAR
    ax.AXIS := Axis;
    ax.OP := 3; ax();
    exEdge := Execute AND NOT exPrev; exPrev := Execute;
    Done := FALSE; CommandAborted := FALSE; Error := FALSE; ErrorID := 0;
    IF NOT active AND exEdge THEN
        IF ModuloFactor <= 0 THEN
            Error := TRUE; ErrorID := 1;
        ELSE
            ax.OP := 4; ax.INDEX := 16#6064; ax();   // pos actual
            // normalize current and target into [0,ModuloFactor)
            cur := ax.VALUE - (ax.VALUE / ModuloFactor) * ModuloFactor;
            IF cur < 0 THEN cur := cur + ModuloFactor; END_IF;
            tgt := Position - (Position / ModuloFactor) * ModuloFactor;
            IF tgt < 0 THEN tgt := tgt + ModuloFactor; END_IF;
            delta := tgt - cur;
            IF Direction = 1 THEN
                IF delta < 0 THEN delta := delta + ModuloFactor; END_IF;
            ELSIF Direction = 2 THEN
                IF delta > 0 THEN delta := delta - ModuloFactor; END_IF;
            ELSE
                IF delta > ModuloFactor / 2 THEN
                    delta := delta - ModuloFactor;
                ELSIF delta < -ModuloFactor / 2 THEN
                    delta := delta + ModuloFactor;
                END_IF;
            END_IF;
            goal := ax.VALUE + delta;
            ax.OP := 5; ax.INDEX := 16#6060; ax.VALUE := 1; ax();
            ax.OP := 5; ax.INDEX := 16#607A; ax.VALUE := goal; ax();
            ax.OP := 5; ax.INDEX := 16#6040; ax.VALUE := 16#001F; ax();
            IF ax.STATUS = 0 THEN
                active := TRUE; rel := TRUE;
            ELSE
                Error := TRUE; ErrorID := ax.ERRID;
            END_IF;
        END_IF;
    ELSIF active THEN
        IF rel THEN
            ax.OP := 5; ax.INDEX := 16#6040; ax.VALUE := 16#000F; ax();
            rel := FALSE;
        END_IF;
        ax.OP := 6; ax();
        IF ax.STATUS < 0 THEN
            Error := TRUE; ErrorID := ax.ERRID; active := FALSE;
        ELSIF ax.TARGET_REACHED = 1 THEN
            Done := TRUE; active := FALSE;
        END_IF;
    END_IF
    Busy := active;
END_FUNCTION_BLOCK

// ---- MC_SetOverride: velocity override factor ----
// While Enable is held the velocity-mode target (0x60FF) is scaled
// to baseVel * VelFactor / 100, where baseVel is latched on the
// Enable rising edge; on release the unscaled base is restored.
// VelFactor is an integer percent (100 = 100%, 0 = hold at rest).
// Applies to velocity modes (PV/VL); ProfilePosition speed comes
// from axis config so the write is a harmless no-op there.
FUNCTION_BLOCK MC_SetOverride
VAR_INPUT
    Enable : BOOL;
    VelFactor : DINT;
    Axis : UDINT;
END_VAR
VAR_OUTPUT
    Enabled : BOOL;
    Busy : BOOL;
END_VAR
VAR
    ax : FB_MotionAxis;
    enPrev : BOOL;
    hasBase : BOOL;
    baseVel : DINT;
END_VAR
    ax.AXIS := Axis;
    ax.OP := 3; ax();
    IF Enable AND NOT enPrev THEN
        ax.OP := 4; ax.INDEX := 16#60FF; ax();
        baseVel := ax.VALUE;
        hasBase := TRUE;
    END_IF;
    enPrev := Enable;
    IF Enable AND hasBase THEN
        ax.OP := 5; ax.INDEX := 16#60FF;
        ax.VALUE := baseVel * VelFactor / 100; ax();
        Enabled := (ax.STATUS = 0);
    ELSIF (NOT Enable) AND hasBase THEN
        ax.OP := 5; ax.INDEX := 16#60FF; ax.VALUE := baseVel; ax();
        hasBase := FALSE;
        Enabled := FALSE;
    ELSE
        Enabled := FALSE;
    END_IF;
    Busy := FALSE;
END_FUNCTION_BLOCK

// ---- MC_ReadParameter: read a DS402 object as an axis parameter ----
// ParameterNumber is the DS402 object index. Valid reports a
// successful read into Value.
FUNCTION_BLOCK MC_ReadParameter
VAR_INPUT
    Enable : BOOL;
    ParameterNumber : UDINT;
    Axis : UDINT;
END_VAR
VAR_OUTPUT
    Valid : BOOL;
    Value : DINT;
    Busy : BOOL;
END_VAR
VAR
    ax : FB_MotionAxis;
END_VAR
    ax.OP := 3; ax();
    ax.AXIS := Axis;
    ax.OP := 4;
    ax.INDEX := ParameterNumber;
    ax();
    IF Enable AND ax.STATUS = 0 THEN
        Valid := TRUE;
        Value := ax.VALUE;
    ELSE
        Valid := FALSE;
        Value := 0;
    END_IF;
    Busy := FALSE;
END_FUNCTION_BLOCK

// ---- MC_WriteParameter: write a DS402 object as an axis parameter ----
// Execute edge writes Value to the object named by ParameterNumber.
FUNCTION_BLOCK MC_WriteParameter
VAR_INPUT
    Execute : BOOL;
    ParameterNumber : UDINT;
    Value : DINT;
    Axis : UDINT;
END_VAR
VAR_OUTPUT
    Done : BOOL;
    Busy : BOOL;
    Error : BOOL;
    ErrorID : UDINT;
END_VAR
VAR
    ax : FB_MotionAxis;
    exPrev : BOOL;
    exEdge : BOOL;
END_VAR
    ax.OP := 3; ax();
    ax.AXIS := Axis;
    exEdge := Execute AND NOT exPrev; exPrev := Execute;
    Done := FALSE; Error := FALSE; ErrorID := 0;
    IF exEdge THEN
        ax.OP := 5;
        ax.INDEX := ParameterNumber;
        ax.VALUE := Value;
        ax();
        IF ax.STATUS = 0 THEN
            Done := TRUE;
        ELSE
            Error := TRUE; ErrorID := ax.ERRID;
        END_IF;
    END_IF;
    Busy := FALSE;
END_FUNCTION_BLOCK

// ---- MC_ReadBoolParameter: read a DS402 object as a BOOL ----
// Value is TRUE when the object at ParameterNumber is nonzero.
FUNCTION_BLOCK MC_ReadBoolParameter
VAR_INPUT
    Enable : BOOL;
    ParameterNumber : UDINT;
    Axis : UDINT;
END_VAR
VAR_OUTPUT
    Valid : BOOL;
    Value : BOOL;
    Busy : BOOL;
END_VAR
VAR
    ax : FB_MotionAxis;
END_VAR
    ax.OP := 3; ax();
    ax.AXIS := Axis;
    ax.OP := 4;
    ax.INDEX := ParameterNumber;
    ax();
    IF Enable AND ax.STATUS = 0 THEN
        Valid := TRUE;
        Value := (ax.VALUE <> 0);
    ELSE
        Valid := FALSE;
        Value := FALSE;
    END_IF;
    Busy := FALSE;
END_FUNCTION_BLOCK

// ---- MC_WriteBoolParameter: write a DS402 object from a BOOL ----
// Execute edge writes 1/0 to the object named by ParameterNumber.
FUNCTION_BLOCK MC_WriteBoolParameter
VAR_INPUT
    Execute : BOOL;
    ParameterNumber : UDINT;
    Value : BOOL;
    Axis : UDINT;
END_VAR
VAR_OUTPUT
    Done : BOOL;
    Busy : BOOL;
    Error : BOOL;
    ErrorID : UDINT;
END_VAR
VAR
    ax : FB_MotionAxis;
    exPrev : BOOL;
    exEdge : BOOL;
    raw : DINT;
END_VAR
    ax.OP := 3; ax();
    ax.AXIS := Axis;
    exEdge := Execute AND NOT exPrev; exPrev := Execute;
    Done := FALSE; Error := FALSE; ErrorID := 0;
    IF exEdge THEN
        IF Value THEN raw := 1; ELSE raw := 0; END_IF;
        ax.OP := 5;
        ax.INDEX := ParameterNumber;
        ax.VALUE := raw;
        ax();
        IF ax.STATUS = 0 THEN
            Done := TRUE;
        ELSE
            Error := TRUE; ErrorID := ax.ERRID;
        END_IF;
    END_IF;
    Busy := FALSE;
END_FUNCTION_BLOCK

// ================================================================== //
// Tranche-5 blocks: touch-probe latch and master/slave gearing.
// MC_TouchProbe captures PositionActualValue on the TriggerInput
// rising edge — a cycle-level software latch (TwinCAT latches in
// drive hardware, sub-cycle; the simulated backend has no latch
// object, so capture latency is one scan — documented gap).
// MC_GearIn couples the slave axis to the master at a velocity
// ratio by reading VelocityActualValue each scan and driving the
// slave's TargetVelocity in PV mode — velocity-ratio coupling, not
// an exact position-phase lock (that needs cyclic setpoint
// coupling / a coupling object; documented gap). MC_AbortTrigger
// cancels an armed probe through the per-axis probe-abort object
// 0x2001 (see below); MC_TouchProbe self-aborts on a re-Execute.
// ================================================================== //

// ---- MC_TouchProbe: position capture on a trigger edge ----
// Execute edge arms the probe. While armed the axis position is
// polled each scan; on a TriggerInput rising edge the position is
// recorded into RecordedPosition (optionally only when inside
// [FirstPosition,LastPosition] when WindowOnly is TRUE). Done
// reports a captured value. Re-executing while armed re-arms.
// The arm edge also clears the axis probe-abort object (0x2001) so
// an abort issued before the arm cannot kill the new cycle; while
// armed each scan polls 0x2001 and a nonzero value consumes the
// request (writes 0 back), disarms and pulses CommandAborted.
FUNCTION_BLOCK MC_TouchProbe
VAR_INPUT
    Execute : BOOL;
    TriggerInput : BOOL;
    WindowOnly : BOOL;
    FirstPosition : DINT;
    LastPosition : DINT;
    Axis : UDINT;
END_VAR
VAR_OUTPUT
    Done : BOOL;
    Busy : BOOL;
    CommandAborted : BOOL;
    Error : BOOL;
    ErrorID : UDINT;
    RecordedPosition : DINT;
END_VAR
VAR
    ax : FB_MotionAxis;
    exPrev : BOOL;
    exEdge : BOOL;
    armed : BOOL;
    trigPrev : BOOL;
    inWin : BOOL;
END_VAR
    ax.AXIS := Axis;
    ax.OP := 3; ax();
    exEdge := Execute AND NOT exPrev; exPrev := Execute;
    Done := FALSE; CommandAborted := FALSE; Error := FALSE; ErrorID := 0;
    IF exEdge THEN
        armed := TRUE;               // (re)arm the probe
        ax.OP := 5; ax.INDEX := 16#2001; ax.VALUE := 0; ax();
    END_IF;
    IF armed THEN
        ax.OP := 4; ax.INDEX := 16#2001; ax();   // abort request?
        IF ax.VALUE <> 0 THEN
            ax.OP := 5; ax.INDEX := 16#2001; ax.VALUE := 0; ax();
            armed := FALSE;
            CommandAborted := TRUE;
        ELSE
            ax.OP := 4; ax.INDEX := 16#6064; ax();   // pos actual
            IF TriggerInput AND NOT trigPrev THEN
                inWin := TRUE;
                IF WindowOnly THEN
                    inWin := (ax.VALUE >= FirstPosition)
                             AND (ax.VALUE <= LastPosition);
                END_IF;
                IF inWin THEN
                    RecordedPosition := ax.VALUE;
                    Done := TRUE;
                    armed := FALSE;
                END_IF;
            END_IF;
        END_IF;
    END_IF;
    trigPrev := TriggerInput;
    Busy := armed;
END_FUNCTION_BLOCK

// ---- MC_AbortTrigger: cancel an armed touch-probe cycle ----
// Execute edge writes 1 to the axis probe-abort object (0x2001,
// manufacturer-specific sim extension shared with MC_TouchProbe).
// Done reports once the request has been consumed, i.e. the flag
// reads 0 again (an armed MC_TouchProbe cleared it after
// disarming). Busy stays TRUE while the request is pending; issue
// aborts only while a probe cycle is active, matching TwinCAT
// usage. TriggerInput is accepted for signature fidelity; the
// single-probe-per-axis model aborts the axis's armed probe
// regardless of which trigger reference is passed.
FUNCTION_BLOCK MC_AbortTrigger
VAR_INPUT
    Execute : BOOL;
    TriggerInput : BOOL;
    Axis : UDINT;
END_VAR
VAR_OUTPUT
    Done : BOOL;
    Busy : BOOL;
    CommandAborted : BOOL;
    Error : BOOL;
    ErrorID : UDINT;
END_VAR
VAR
    ax : FB_MotionAxis;
    exPrev : BOOL;
    exEdge : BOOL;
    pending : BOOL;
END_VAR
    ax.AXIS := Axis;
    ax.OP := 3; ax();
    exEdge := Execute AND NOT exPrev; exPrev := Execute;
    Done := FALSE; Busy := pending; CommandAborted := FALSE;
    Error := FALSE; ErrorID := 0;
    IF exEdge AND NOT pending THEN
        ax.OP := 5; ax.INDEX := 16#2001; ax.VALUE := 1; ax();
        IF ax.STATUS = 0 THEN
            pending := TRUE;
        ELSE
            Error := TRUE; ErrorID := ax.ERRID;
        END_IF;
    END_IF;
    IF pending THEN
        ax.OP := 4; ax.INDEX := 16#2001; ax();
        IF ax.STATUS = 0 AND ax.VALUE = 0 THEN
            Done := TRUE; pending := FALSE;
        END_IF;
    END_IF;
    Busy := pending;
END_FUNCTION_BLOCK

// ---- MC_GearIn: velocity-ratio master/slave coupling ----
// While Execute is held the slave axis runs in ProfileVelocity at
// TargetVelocity = master VelocityActualValue * RatioNumerator /
// RatioDenominator, so the slave velocity tracks the master at the
// gear ratio (positions track proportionally but not phase-locked).
// Engage edge puts the slave into PV mode + enable; on release the
// slave keeps its last velocity until MC_GearOut/MC_Halt stops it.
FUNCTION_BLOCK MC_GearIn
VAR_INPUT
    Execute : BOOL;
    RatioNumerator : DINT;
    RatioDenominator : DINT;
    Acceleration : DINT;
    Deceleration : DINT;
    Master : UDINT;
    Slave : UDINT;
END_VAR
VAR_OUTPUT
    InGear : BOOL;
    Busy : BOOL;
    CommandAborted : BOOL;
    Error : BOOL;
    ErrorID : UDINT;
END_VAR
VAR
    axM : FB_MotionAxis;
    axS : FB_MotionAxis;
    exPrev : BOOL;
    exEdge : BOOL;
    mvel : DINT;
END_VAR
    axM.AXIS := Master;
    axS.AXIS := Slave;
    axM.OP := 3; axM();
    exEdge := Execute AND NOT exPrev; exPrev := Execute;
    InGear := FALSE; CommandAborted := FALSE; Error := FALSE; ErrorID := 0;
    IF exEdge THEN
        IF RatioDenominator = 0 THEN
            Error := TRUE; ErrorID := 1;
        ELSE
            axS.OP := 5; axS.INDEX := 16#6040; axS.VALUE := 16#000F; axS();
            axS.OP := 5; axS.INDEX := 16#6060; axS.VALUE := 3; axS();
        END_IF;
    END_IF;
    IF Execute AND RatioDenominator <> 0 THEN
        // slave velocity follows the master at the gear ratio
        axM.OP := 4; axM.INDEX := 16#606C; axM();
        mvel := axM.VALUE;
        axS.OP := 5; axS.INDEX := 16#60FF;
        axS.VALUE := mvel * RatioNumerator / RatioDenominator; axS();
        axS.OP := 6; axS();
        IF axS.STATUS < 0 THEN
            Error := TRUE; ErrorID := axS.ERRID;
        ELSE
            InGear := TRUE;
        END_IF;
    END_IF;
    Busy := Execute AND (RatioDenominator <> 0);
END_FUNCTION_BLOCK

// ---- MC_GearOut: uncouple the slave and ramp it to rest ----
// Execute edge commands the slave TargetVelocity to 0 (PV decel);
// Done when VelocityActualValue reaches zero. The slave stays
// enabled in velocity mode; use MC_Halt/MC_Stop for a hard stop.
FUNCTION_BLOCK MC_GearOut
VAR_INPUT
    Execute : BOOL;
    Deceleration : DINT;
    Slave : UDINT;
END_VAR
VAR_OUTPUT
    Done : BOOL;
    Busy : BOOL;
    Error : BOOL;
    ErrorID : UDINT;
END_VAR
VAR
    axS : FB_MotionAxis;
    exPrev : BOOL;
    exEdge : BOOL;
    active : BOOL;
END_VAR
    axS.AXIS := Slave;
    axS.OP := 3; axS();
    exEdge := Execute AND NOT exPrev; exPrev := Execute;
    Done := FALSE; Error := FALSE; ErrorID := 0;
    IF NOT active AND exEdge THEN
        axS.OP := 5; axS.INDEX := 16#60FF; axS.VALUE := 0; axS();
        active := TRUE;
    ELSIF active THEN
        axS.OP := 6; axS();
        IF axS.STATUS < 0 THEN
            Error := TRUE; ErrorID := axS.ERRID; active := FALSE;
        ELSIF axS.VEL_ACTUAL = 0 THEN
            Done := TRUE; active := FALSE;
        END_IF;
    END_IF;
    Busy := active;
END_FUNCTION_BLOCK
